Universal Robots URScript: FaiChun_9 Jan_5.script

def Machining1():
  # Default parameters:
  global speed_ms = 0.03
  global speed_rads = 0.75
  global accel_mss = 3
  global accel_radss = 1.2
  global blend_radius_m = 0.0003

  # Add subprograms here
  # Start of main program
  # Program generated by RoboDK v5.6.8 for UR10e on 09/01/2025 17:26:35
  # Using nominal kinematics.
  blend_radius_m = 0.0003
  speed_ms = 0.03
  # set_reference(p[0.325000, -0.070000, 0.000000, 0.000000, 0.000000, 0.000000])
  set_tcp(p[0.000000, 0.000000, 0.252000, 0.000000, 0.000000, 0.000000])
  # Show Tool
  movej([0.354568, -1.073416, -2.632395, -1.006578, 1.570796, 1.925364],accel_radss,speed_rads,0,blend_radius_m)
  movel([0.354568, -1.133460, -2.672124, -0.906805, 1.570796, 1.925364],accel_mss,speed_ms,0,blend_radius_m)
  #SetTool1
  #M_RunCode6
  #3SetRPM60000
  speed_ms = 0.03
  #M_RunCode3
  movel([0.354568, -1.161287, -2.687269, -0.863833, 1.570796, 1.925364],accel_mss,speed_ms,0,blend_radius_m)
  speed_ms = 0.003
  movel([0.354568, -1.168634, -2.690994, -0.852761, 1.570796, 1.925364],accel_mss,speed_ms,0,blend_radius_m)
  speed_ms = 0.007
  movel([0.356966, -1.171496, -2.689722, -0.851171, 1.570796, 1.927762],accel_mss,speed_ms,0,blend_radius_m)
  movel([0.359544, -1.173577, -2.688792, -0.850019, 1.570796, 1.930340],accel_mss,speed_ms,0,blend_radius_m)
  movel([0.362316, -1.174874, -2.688211, -0.849304, 1.570796, 1.933112],accel_mss,speed_ms,0,blend_radius_m)
  movel([0.365281, -1.175393, -2.687978, -0.849019, 1.570796, 1.936077],accel_mss,speed_ms,0,blend_radius_m)
  movel([0.368380, -1.175227, -2.688052, -0.849110, 1.570796, 1.939176],accel_mss,speed_ms,0,blend_radius_m)
  movel([0.371545, -1.174464, -2.688395, -0.849530, 1.570796, 1.942341],accel_mss,speed_ms,0,blend_radius_m)
  movel([0.374787, -1.173102, -2.689005, -0.850282, 1.570796, 1.945583],accel_mss,speed_ms,0,blend_radius_m)
  movel([0.378111, -1.171130, -2.689885, -0.851373, 1.570796, 1.948907],accel_mss,speed_ms,0,blend_radius_m)
  movel([0.363017, -1.184266, -2.683945, -0.844178, 1.570796, 1.933813],accel_mss,speed_ms,0,blend_radius_m)
  movel([0.342026, -1.154782, -2.697027, -0.860579, 1.570796, 1.912822],accel_mss,speed_ms,0,blend_radius_m)
  movel([0.343555, -1.153375, -2.697629, -0.861384, 1.570796, 1.914352],accel_mss,speed_ms,0,blend_radius_m)
  movel([0.347706, -1.150135, -2.699008, -0.863246, 1.570796, 1.918503],accel_mss,speed_ms,0,blend_radius_m)
  movel([0.352300, -1.147640, -2.700062, -0.864686, 1.570796, 1.923096],accel_mss,speed_ms,0,blend_radius_m)
  movel([0.357069, -1.145805, -2.700834, -0.865750, 1.570796, 1.927865],accel_mss,speed_ms,0,blend_radius_m)
  movel([0.361749, -1.144532, -2.701367, -0.866490, 1.570796, 1.932545],accel_mss,speed_ms,0,blend_radius_m)
  movel([0.373963, -1.142426, -2.702246, -0.867717, 1.570796, 1.944759],accel_mss,speed_ms,0,blend_radius_m)
  movel([0.385222, -1.140714, -2.702957, -0.868719, 1.570796, 1.956018],accel_mss,speed_ms,0,blend_radius_m)
  movel([0.389576, -1.139664, -2.703391, -0.869334, 1.570796, 1.960373],accel_mss,speed_ms,0,blend_radius_m)
  movel([0.393934, -1.138139, -2.704021, -0.870229, 1.570796, 1.964730],accel_mss,speed_ms,0,blend_radius_m)
  movel([0.398079, -1.136054, -2.704878, -0.871458, 1.570796, 1.968876],accel_mss,speed_ms,0,blend_radius_m)
  movel([0.401806, -1.133312, -2.705998, -0.873079, 1.570796, 1.972603],accel_mss,speed_ms,0,blend_radius_m)
  movel([0.405715, -1.129228, -2.707653, -0.875508, 1.570796, 1.976512],accel_mss,speed_ms,0,blend_radius_m)
  movel([0.407057, -1.127215, -2.708462, -0.876712, 1.570796, 1.977853],accel_mss,speed_ms,0,blend_radius_m)
  movel([0.407988, -1.125220, -2.709261, -0.877908, 1.570796, 1.978784],accel_mss,speed_ms,0,blend_radius_m)
  movel([0.408720, -1.121628, -2.710690, -0.880072, 1.570796, 1.979516],accel_mss,speed_ms,0,blend_radius_m)
  movel([0.408019, -1.118804, -2.711804, -0.881781, 1.570796, 1.978816],accel_mss,speed_ms,0,blend_radius_m)
  movel([0.406875, -1.117482, -2.712323, -0.882584, 1.570796, 1.977671],accel_mss,speed_ms,0,blend_radius_m)
  movel([0.405474, -1.116991, -2.712516, -0.882883, 1.570796, 1.976271],accel_mss,speed_ms,0,blend_radius_m)
  movel([0.403971, -1.117249, -2.712414, -0.882726, 1.570796, 1.974768],accel_mss,speed_ms,0,blend_radius_m)
  movel([0.402512, -1.118181, -2.712049, -0.882159, 1.570796, 1.973309],accel_mss,speed_ms,0,blend_radius_m)
  movel([0.400903, -1.120447, -2.711157, -0.880785, 1.570796, 1.971699],accel_mss,speed_ms,0,blend_radius_m)
  movel([0.399463, -1.122720, -2.710257, -0.879412, 1.570796, 1.970259],accel_mss,speed_ms,0,blend_radius_m)
  movel([0.397172, -1.125110, -2.709305, -0.877974, 1.570796, 1.967968],accel_mss,speed_ms,0,blend_radius_m)
  movel([0.394069, -1.127271, -2.708440, -0.876678, 1.570796, 1.964865],accel_mss,speed_ms,0,blend_radius_m)
  movel([0.391233, -1.128021, -2.708139, -0.876230, 1.570796, 1.962029],accel_mss,speed_ms,0,blend_radius_m)
  movel([0.388876, -1.127540, -2.708332, -0.876517, 1.570796, 1.959673],accel_mss,speed_ms,0,blend_radius_m)
  movel([0.387215, -1.125994, -2.708952, -0.877443, 1.570796, 1.958012],accel_mss,speed_ms,0,blend_radius_m)
  movel([0.386430, -1.123660, -2.709883, -0.878846, 1.570796, 1.957226],accel_mss,speed_ms,0,blend_radius_m)
  movel([0.386711, -1.120809, -2.711013, -0.880566, 1.570796, 1.957507],accel_mss,speed_ms,0,blend_radius_m)
  movel([0.388136, -1.117739, -2.712222, -0.882428, 1.570796, 1.958932],accel_mss,speed_ms,0,blend_radius_m)
  movel([0.390789, -1.114754, -2.713389, -0.884246, 1.570796, 1.961586],accel_mss,speed_ms,0,blend_radius_m)
  movel([0.393483, -1.112681, -2.714194, -0.885514, 1.570796, 1.964280],accel_mss,speed_ms,0,blend_radius_m)
  movel([0.396144, -1.111333, -2.714716, -0.886340, 1.570796, 1.966940],accel_mss,speed_ms,0,blend_radius_m)
  movel([0.398770, -1.110715, -2.714954, -0.886719, 1.570796, 1.969567],accel_mss,speed_ms,0,blend_radius_m)
  movel([0.401345, -1.110843, -2.714905, -0.886641, 1.570796, 1.972141],accel_mss,speed_ms,0,blend_radius_m)
  movel([0.403780, -1.111624, -2.714603, -0.886161, 1.570796, 1.974576],accel_mss,speed_ms,0,blend_radius_m)
  movel([0.405978, -1.112973, -2.714081, -0.885335, 1.570796, 1.976774],accel_mss,speed_ms,0,blend_radius_m)
  movel([0.409660, -1.117365, -2.712369, -0.882655, 1.570796, 1.980457],accel_mss,speed_ms,0,blend_radius_m)
  movel([0.411296, -1.120837, -2.711002, -0.880549, 1.570796, 1.982092],accel_mss,speed_ms,0,blend_radius_m)
  movel([0.412317, -1.124558, -2.709525, -0.878306, 1.570796, 1.983113],accel_mss,speed_ms,0,blend_radius_m)
  movel([0.412731, -1.128520, -2.707938, -0.875931, 1.570796, 1.983527],accel_mss,speed_ms,0,blend_radius_m)
  movel([0.412549, -1.132708, -2.706243, -0.873438, 1.570796, 1.983345],accel_mss,speed_ms,0,blend_radius_m)
  movel([0.411547, -1.136963, -2.704504, -0.870921, 1.570796, 1.982343],accel_mss,speed_ms,0,blend_radius_m)
  movel([0.409511, -1.141125, -2.702786, -0.868478, 1.570796, 1.980307],accel_mss,speed_ms,0,blend_radius_m)
  movel([0.406444, -1.145198, -2.701088, -0.866103, 1.570796, 1.977240],accel_mss,speed_ms,0,blend_radius_m)
  movel([0.402358, -1.149188, -2.699409, -0.863792, 1.570796, 1.973154],accel_mss,speed_ms,0,blend_radius_m)
  movel([0.398284, -1.152264, -2.698104, -0.862022, 1.570796, 1.969081],accel_mss,speed_ms,0,blend_radius_m)
  movel([0.394157, -1.154540, -2.697131, -0.860718, 1.570796, 1.964954],accel_mss,speed_ms,0,blend_radius_m)
  movel([0.390077, -1.156158, -2.696437, -0.859794, 1.570796, 1.960874],accel_mss,speed_ms,0,blend_radius_m)
  movel([0.386157, -1.157252, -2.695966, -0.859171, 1.570796, 1.956954],accel_mss,speed_ms,0,blend_radius_m)
  movel([0.376830, -1.158761, -2.695314, -0.858314, 1.570796, 1.947626],accel_mss,speed_ms,0,blend_radius_m)
  movel([0.367992, -1.160305, -2.694646, -0.857439, 1.570796, 1.938788],accel_mss,speed_ms,0,blend_radius_m)
  movel([0.364425, -1.161338, -2.694196, -0.856855, 1.570796, 1.935222],accel_mss,speed_ms,0,blend_radius_m)
  movel([0.360783, -1.162831, -2.693545, -0.856012, 1.570796, 1.931580],accel_mss,speed_ms,0,blend_radius_m)
  movel([0.357192, -1.164865, -2.692655, -0.854869, 1.570796, 1.927988],accel_mss,speed_ms,0,blend_radius_m)
  movel([0.353786, -1.167525, -2.691484, -0.853380, 1.570796, 1.924582],accel_mss,speed_ms,0,blend_radius_m)
  movel([0.354568, -1.168634, -2.690994, -0.852761, 1.570796, 1.925364],accel_mss,speed_ms,0,blend_radius_m)
  speed_ms = 0.003
  movel([0.354568, -1.161287, -2.687269, -0.863833, 1.570796, 1.925364],accel_mss,speed_ms,0,blend_radius_m)
  speed_ms = 0.03
  movel([0.354568, -1.133460, -2.672124, -0.906805, 1.570796, 1.925364],accel_mss,speed_ms,0,blend_radius_m)
  #M_RunCode9
  movel([0.379678, -1.157713, -2.661566, -0.893110, 1.570796, 1.950474],accel_mss,speed_ms,0,blend_radius_m)
  #M_RunCode3
  movel([0.379678, -1.185401, -2.676392, -0.850596, 1.570796, 1.950474],accel_mss,speed_ms,0,blend_radius_m)
  speed_ms = 0.003
  movel([0.379678, -1.192696, -2.680036, -0.839657, 1.570796, 1.950474],accel_mss,speed_ms,0,blend_radius_m)
  speed_ms = 0.007
  movel([0.387460, -1.185010, -2.683603, -0.843776, 1.570796, 1.958256],accel_mss,speed_ms,0,blend_radius_m)
  movel([0.399155, -1.174764, -2.688260, -0.849365, 1.570796, 1.969951],accel_mss,speed_ms,0,blend_radius_m)
  movel([0.411336, -1.164890, -2.692644, -0.854855, 1.570796, 1.982132],accel_mss,speed_ms,0,blend_radius_m)
  movel([0.420366, -1.158451, -2.695449, -0.858490, 1.570796, 1.991162],accel_mss,speed_ms,0,blend_radius_m)
  movel([0.423713, -1.156585, -2.696253, -0.859551, 1.570796, 1.994510],accel_mss,speed_ms,0,blend_radius_m)
  movel([0.426343, -1.155682, -2.696642, -0.860066, 1.570796, 1.997139],accel_mss,speed_ms,0,blend_radius_m)
  movel([0.428246, -1.155744, -2.696615, -0.860030, 1.570796, 1.999042],accel_mss,speed_ms,0,blend_radius_m)
  movel([0.429420, -1.156775, -2.696172, -0.859443, 1.570796, 2.000216],accel_mss,speed_ms,0,blend_radius_m)
  movel([0.429733, -1.158510, -2.695423, -0.858456, 1.570796, 2.000529],accel_mss,speed_ms,0,blend_radius_m)
  movel([0.429055, -1.160703, -2.694472, -0.857213, 1.570796, 1.999851],accel_mss,speed_ms,0,blend_radius_m)
  movel([0.427394, -1.163343, -2.693322, -0.855724, 1.570796, 1.998190],accel_mss,speed_ms,0,blend_radius_m)
  movel([0.424759, -1.166426, -2.691969, -0.853994, 1.570796, 1.995555],accel_mss,speed_ms,0,blend_radius_m)
  movel([0.416644, -1.174214, -2.688507, -0.849668, 1.570796, 1.987440],accel_mss,speed_ms,0,blend_radius_m)
  movel([0.404851, -1.184338, -2.683912, -0.844139, 1.570796, 1.975647],accel_mss,speed_ms,0,blend_radius_m)
  movel([0.392963, -1.193873, -2.679484, -0.839032, 1.570796, 1.963760],accel_mss,speed_ms,0,blend_radius_m)
  movel([0.384351, -1.200009, -2.676582, -0.835798, 1.570796, 1.955147],accel_mss,speed_ms,0,blend_radius_m)
  movel([0.381176, -1.201791, -2.675731, -0.834866, 1.570796, 1.951973],accel_mss,speed_ms,0,blend_radius_m)
  movel([0.378665, -1.202681, -2.675305, -0.834403, 1.570796, 1.949461],accel_mss,speed_ms,0,blend_radius_m)
  movel([0.376810, -1.202676, -2.675308, -0.834405, 1.570796, 1.947607],accel_mss,speed_ms,0,blend_radius_m)
  movel([0.375605, -1.201780, -2.675737, -0.834872, 1.570796, 1.946401],accel_mss,speed_ms,0,blend_radius_m)
  movel([0.375198, -1.200206, -2.676488, -0.835695, 1.570796, 1.945994],accel_mss,speed_ms,0,blend_radius_m)
  movel([0.375736, -1.198170, -2.677456, -0.836763, 1.570796, 1.946532],accel_mss,speed_ms,0,blend_radius_m)
  movel([0.377227, -1.195668, -2.678639, -0.838082, 1.570796, 1.948024],accel_mss,speed_ms,0,blend_radius_m)
  movel([0.379678, -1.192696, -2.680036, -0.839657, 1.570796, 1.950474],accel_mss,speed_ms,0,blend_radius_m)
  speed_ms = 0.003
  movel([0.379678, -1.185401, -2.676392, -0.850596, 1.570796, 1.950474],accel_mss,speed_ms,0,blend_radius_m)
  speed_ms = 0.03
  movel([0.379678, -1.157713, -2.661566, -0.893110, 1.570796, 1.950474],accel_mss,speed_ms,0,blend_radius_m)
  #M_RunCode9
  movel([0.372229, -1.160949, -2.660112, -0.891327, 1.570796, 1.943026],accel_mss,speed_ms,0,blend_radius_m)
  #M_RunCode3
  movel([0.372229, -1.188615, -2.674896, -0.848878, 1.570796, 1.943026],accel_mss,speed_ms,0,blend_radius_m)
  speed_ms = 0.003
  movel([0.372229, -1.195902, -2.678528, -0.837958, 1.570796, 1.943026],accel_mss,speed_ms,0,blend_radius_m)
  speed_ms = 0.007
  movel([0.372519, -1.193032, -2.679878, -0.839479, 1.570796, 1.943316],accel_mss,speed_ms,0,blend_radius_m)
  movel([0.373292, -1.189945, -2.681319, -0.841124, 1.570796, 1.944089],accel_mss,speed_ms,0,blend_radius_m)
  movel([0.374568, -1.186684, -2.682831, -0.842874, 1.570796, 1.945364],accel_mss,speed_ms,0,blend_radius_m)
  movel([0.376355, -1.183240, -2.684415, -0.844734, 1.570796, 1.947151],accel_mss,speed_ms,0,blend_radius_m)
  movel([0.378653, -1.179619, -2.686067, -0.846703, 1.570796, 1.949450],accel_mss,speed_ms,0,blend_radius_m)
  movel([0.381456, -1.175876, -2.687760, -0.848753, 1.570796, 1.952252],accel_mss,speed_ms,0,blend_radius_m)
  movel([0.384749, -1.172089, -2.689458, -0.850842, 1.570796, 1.955546],accel_mss,speed_ms,0,blend_radius_m)
  movel([0.388543, -1.168254, -2.691162, -0.852973, 1.570796, 1.959339],accel_mss,speed_ms,0,blend_radius_m)
  movel([0.392836, -1.164375, -2.692870, -0.855144, 1.570796, 1.963633],accel_mss,speed_ms,0,blend_radius_m)
  movel([0.397312, -1.160734, -2.694459, -0.857196, 1.570796, 1.968109],accel_mss,speed_ms,0,blend_radius_m)
  movel([0.401640, -1.157615, -2.695810, -0.858965, 1.570796, 1.972436],accel_mss,speed_ms,0,blend_radius_m)
  movel([0.405819, -1.155020, -2.696926, -0.860443, 1.570796, 1.976615],accel_mss,speed_ms,0,blend_radius_m)
  movel([0.409833, -1.152965, -2.697805, -0.861619, 1.570796, 1.980629],accel_mss,speed_ms,0,blend_radius_m)
  movel([0.413614, -1.151451, -2.698450, -0.862489, 1.570796, 1.984410],accel_mss,speed_ms,0,blend_radius_m)
  movel([0.417092, -1.150479, -2.698862, -0.863048, 1.570796, 1.987889],accel_mss,speed_ms,0,blend_radius_m)
  movel([0.420254, -1.150059, -2.699040, -0.863290, 1.570796, 1.991051],accel_mss,speed_ms,0,blend_radius_m)
  movel([0.423104, -1.150185, -2.698987, -0.863217, 1.570796, 1.993900],accel_mss,speed_ms,0,blend_radius_m)
  movel([0.425609, -1.150820, -2.698717, -0.862851, 1.570796, 1.996406],accel_mss,speed_ms,0,blend_radius_m)
  movel([0.427747, -1.151930, -2.698246, -0.862214, 1.570796, 1.998543],accel_mss,speed_ms,0,blend_radius_m)
  movel([0.429513, -1.153503, -2.697575, -0.861311, 1.570796, 2.000309],accel_mss,speed_ms,0,blend_radius_m)
  movel([0.430906, -1.155546, -2.696700, -0.860143, 1.570796, 2.001703],accel_mss,speed_ms,0,blend_radius_m)
  movel([0.431874, -1.157931, -2.695673, -0.858785, 1.570796, 2.002670],accel_mss,speed_ms,0,blend_radius_m)
  movel([0.432358, -1.160544, -2.694541, -0.857303, 1.570796, 2.003155],accel_mss,speed_ms,0,blend_radius_m)
  movel([0.432364, -1.163381, -2.693305, -0.855703, 1.570796, 2.003160],accel_mss,speed_ms,0,blend_radius_m)
  movel([0.431892, -1.166435, -2.691965, -0.853989, 1.570796, 2.002688],accel_mss,speed_ms,0,blend_radius_m)
  movel([0.430933, -1.169665, -2.690537, -0.852187, 1.570796, 2.001729],accel_mss,speed_ms,0,blend_radius_m)
  movel([0.429473, -1.173023, -2.689040, -0.850325, 1.570796, 2.000269],accel_mss,speed_ms,0,blend_radius_m)
  movel([0.427521, -1.176505, -2.687476, -0.848407, 1.570796, 1.998318],accel_mss,speed_ms,0,blend_radius_m)
  movel([0.425078, -1.180116, -2.685842, -0.846432, 1.570796, 1.995874],accel_mss,speed_ms,0,blend_radius_m)
  movel([0.422172, -1.183774, -2.684170, -0.844444, 1.570796, 1.992968],accel_mss,speed_ms,0,blend_radius_m)
  movel([0.418832, -1.187414, -2.682494, -0.842481, 1.570796, 1.989629],accel_mss,speed_ms,0,blend_radius_m)
  movel([0.415055, -1.191041, -2.680809, -0.840539, 1.570796, 1.985852],accel_mss,speed_ms,0,blend_radius_m)
  movel([0.410849, -1.194652, -2.679117, -0.838619, 1.570796, 1.981646],accel_mss,speed_ms,0,blend_radius_m)
  movel([0.406521, -1.198006, -2.677534, -0.836850, 1.570796, 1.977317],accel_mss,speed_ms,0,blend_radius_m)
  movel([0.402383, -1.200845, -2.676183, -0.835360, 1.570796, 1.973179],accel_mss,speed_ms,0,blend_radius_m)
  movel([0.398419, -1.203189, -2.675062, -0.834138, 1.570796, 1.969215],accel_mss,speed_ms,0,blend_radius_m)
  movel([0.394629, -1.205036, -2.674174, -0.833179, 1.570796, 1.965426],accel_mss,speed_ms,0,blend_radius_m)
  movel([0.391062, -1.206401, -2.673515, -0.832473, 1.570796, 1.961858],accel_mss,speed_ms,0,blend_radius_m)
  movel([0.387772, -1.207286, -2.673087, -0.832016, 1.570796, 1.958568],accel_mss,speed_ms,0,blend_radius_m)
  movel([0.384754, -1.207698, -2.672887, -0.831804, 1.570796, 1.955550],accel_mss,speed_ms,0,blend_radius_m)
  movel([0.382004, -1.207633, -2.672919, -0.831838, 1.570796, 1.952800],accel_mss,speed_ms,0,blend_radius_m)
  movel([0.379552, -1.207117, -2.673169, -0.832104, 1.570796, 1.950348],accel_mss,speed_ms,0,blend_radius_m)
  movel([0.377425, -1.206179, -2.673622, -0.832588, 1.570796, 1.948222],accel_mss,speed_ms,0,blend_radius_m)
  movel([0.375621, -1.204815, -2.674280, -0.833294, 1.570796, 1.946417],accel_mss,speed_ms,0,blend_radius_m)
  movel([0.374138, -1.203022, -2.675142, -0.834225, 1.570796, 1.944934],accel_mss,speed_ms,0,blend_radius_m)
  movel([0.373043, -1.200893, -2.676161, -0.835336, 1.570796, 1.943839],accel_mss,speed_ms,0,blend_radius_m)
  movel([0.372405, -1.198522, -2.677289, -0.836578, 1.570796, 1.943201],accel_mss,speed_ms,0,blend_radius_m)
  movel([0.372229, -1.195902, -2.678528, -0.837958, 1.570796, 1.943026],accel_mss,speed_ms,0,blend_radius_m)
  speed_ms = 0.003
  movel([0.372229, -1.188615, -2.674896, -0.848878, 1.570796, 1.943026],accel_mss,speed_ms,0,blend_radius_m)
  speed_ms = 0.03
  movel([0.372229, -1.160949, -2.660112, -0.891327, 1.570796, 1.943026],accel_mss,speed_ms,0,blend_radius_m)
  #M_RunCode9
  movel([0.502532, -1.419663, -2.504293, -0.788433, 1.570796, 2.073328],accel_mss,speed_ms,0,blend_radius_m)
  #M_RunCode3
  movel([0.502532, -1.443463, -2.515724, -0.753202, 1.570796, 2.073328],accel_mss,speed_ms,0,blend_radius_m)
  speed_ms = 0.003
  movel([0.502532, -1.449619, -2.518509, -0.744260, 1.570796, 2.073328],accel_mss,speed_ms,0,blend_radius_m)
  speed_ms = 0.007
  movel([0.503681, -1.448967, -2.519037, -0.744386, 1.570796, 2.074477],accel_mss,speed_ms,0,blend_radius_m)
  movel([0.506715, -1.447598, -2.520141, -0.744650, 1.570796, 2.077511],accel_mss,speed_ms,0,blend_radius_m)
  movel([0.509926, -1.446841, -2.520750, -0.744798, 1.570796, 2.080722],accel_mss,speed_ms,0,blend_radius_m)
  movel([0.513159, -1.446571, -2.520967, -0.744851, 1.570796, 2.083955],accel_mss,speed_ms,0,blend_radius_m)
  movel([0.516261, -1.446673, -2.520885, -0.744831, 1.570796, 2.087058],accel_mss,speed_ms,0,blend_radius_m)
  movel([0.524203, -1.447750, -2.520018, -0.744621, 1.570796, 2.094999],accel_mss,speed_ms,0,blend_radius_m)
  movel([0.531487, -1.448876, -2.519110, -0.744403, 1.570796, 2.102283],accel_mss,speed_ms,0,blend_radius_m)
  movel([0.534346, -1.449044, -2.518974, -0.744371, 1.570796, 2.105142],accel_mss,speed_ms,0,blend_radius_m)
  movel([0.537257, -1.448890, -2.519099, -0.744400, 1.570796, 2.108054],accel_mss,speed_ms,0,blend_radius_m)
  movel([0.540096, -1.448313, -2.519564, -0.744512, 1.570796, 2.110892],accel_mss,speed_ms,0,blend_radius_m)
  movel([0.542736, -1.447217, -2.520447, -0.744724, 1.570796, 2.113533],accel_mss,speed_ms,0,blend_radius_m)
  movel([0.545632, -1.445261, -2.522019, -0.745109, 1.570796, 2.116429],accel_mss,speed_ms,0,blend_radius_m)
  movel([0.546690, -1.444183, -2.522883, -0.745323, 1.570796, 2.117486],accel_mss,speed_ms,0,blend_radius_m)
  movel([0.547489, -1.443035, -2.523801, -0.745553, 1.570796, 2.118285],accel_mss,speed_ms,0,blend_radius_m)
  movel([0.548333, -1.440787, -2.525592, -0.746010, 1.570796, 2.119129],accel_mss,speed_ms,0,blend_radius_m)
  movel([0.548201, -1.438765, -2.527197, -0.746427, 1.570796, 2.118997],accel_mss,speed_ms,0,blend_radius_m)
  movel([0.547632, -1.437654, -2.528076, -0.746659, 1.570796, 2.118428],accel_mss,speed_ms,0,blend_radius_m)
  movel([0.546815, -1.437041, -2.528560, -0.746788, 1.570796, 2.117611],accel_mss,speed_ms,0,blend_radius_m)
  movel([0.545850, -1.436910, -2.528664, -0.746815, 1.570796, 2.116646],accel_mss,speed_ms,0,blend_radius_m)
  movel([0.544842, -1.437235, -2.528407, -0.746747, 1.570796, 2.115638],accel_mss,speed_ms,0,blend_radius_m)
  movel([0.543588, -1.438420, -2.527470, -0.746499, 1.570796, 2.114384],accel_mss,speed_ms,0,blend_radius_m)
  movel([0.542440, -1.439645, -2.526499, -0.746245, 1.570796, 2.113236],accel_mss,speed_ms,0,blend_radius_m)
  movel([0.540743, -1.440783, -2.525595, -0.746011, 1.570796, 2.111539],accel_mss,speed_ms,0,blend_radius_m)
  movel([0.538563, -1.441600, -2.524945, -0.745844, 1.570796, 2.109360],accel_mss,speed_ms,0,blend_radius_m)
  movel([0.536708, -1.441527, -2.525003, -0.745859, 1.570796, 2.107504],accel_mss,speed_ms,0,blend_radius_m)
  movel([0.535289, -1.440723, -2.525643, -0.746023, 1.570796, 2.106086],accel_mss,speed_ms,0,blend_radius_m)
  movel([0.534426, -1.439342, -2.526740, -0.746307, 1.570796, 2.105222],accel_mss,speed_ms,0,blend_radius_m)
  movel([0.534206, -1.437610, -2.528111, -0.746668, 1.570796, 2.105002],accel_mss,speed_ms,0,blend_radius_m)
  movel([0.534705, -1.435753, -2.529576, -0.747060, 1.570796, 2.105502],accel_mss,speed_ms,0,blend_radius_m)
  movel([0.535944, -1.433987, -2.530964, -0.747438, 1.570796, 2.106741],accel_mss,speed_ms,0,blend_radius_m)
  movel([0.537934, -1.432538, -2.532100, -0.747751, 1.570796, 2.108730],accel_mss,speed_ms,0,blend_radius_m)
  movel([0.539842, -1.431708, -2.532749, -0.747932, 1.570796, 2.110639],accel_mss,speed_ms,0,blend_radius_m)
  movel([0.541646, -1.431359, -2.533022, -0.748008, 1.570796, 2.112443],accel_mss,speed_ms,0,blend_radius_m)
  movel([0.543341, -1.431492, -2.532918, -0.747979, 1.570796, 2.114137],accel_mss,speed_ms,0,blend_radius_m)
  movel([0.544925, -1.432107, -2.532437, -0.747845, 1.570796, 2.115721],accel_mss,speed_ms,0,blend_radius_m)
  movel([0.546349, -1.433124, -2.531641, -0.747624, 1.570796, 2.117145],accel_mss,speed_ms,0,blend_radius_m)
  movel([0.547567, -1.434472, -2.530584, -0.747334, 1.570796, 2.118363],accel_mss,speed_ms,0,blend_radius_m)
  movel([0.549380, -1.438137, -2.527694, -0.746558, 1.570796, 2.120176],accel_mss,speed_ms,0,blend_radius_m)
  movel([0.550024, -1.440778, -2.525599, -0.746012, 1.570796, 2.120821],accel_mss,speed_ms,0,blend_radius_m)
  movel([0.550264, -1.443459, -2.523462, -0.745468, 1.570796, 2.121061],accel_mss,speed_ms,0,blend_radius_m)
  movel([0.550102, -1.446181, -2.521280, -0.744927, 1.570796, 2.120899],accel_mss,speed_ms,0,blend_radius_m)
  movel([0.549541, -1.448944, -2.519055, -0.744390, 1.570796, 2.120337],accel_mss,speed_ms,0,blend_radius_m)
  movel([0.548461, -1.451593, -2.516910, -0.743886, 1.570796, 2.119258],accel_mss,speed_ms,0,blend_radius_m)
  movel([0.546732, -1.453987, -2.514963, -0.743439, 1.570796, 2.117528],accel_mss,speed_ms,0,blend_radius_m)
  movel([0.544360, -1.456125, -2.513216, -0.743048, 1.570796, 2.115156],accel_mss,speed_ms,0,blend_radius_m)
  movel([0.541346, -1.458015, -2.511666, -0.742708, 1.570796, 2.112142],accel_mss,speed_ms,0,blend_radius_m)
  movel([0.538430, -1.459300, -2.510609, -0.742480, 1.570796, 2.109226],accel_mss,speed_ms,0,blend_radius_m)
  movel([0.535563, -1.460034, -2.510004, -0.742351, 1.570796, 2.106359],accel_mss,speed_ms,0,blend_radius_m)
  movel([0.532795, -1.460332, -2.509758, -0.742299, 1.570796, 2.103591],accel_mss,speed_ms,0,blend_radius_m)
  movel([0.530186, -1.460301, -2.509784, -0.742304, 1.570796, 2.100982],accel_mss,speed_ms,0,blend_radius_m)
  movel([0.524093, -1.459478, -2.510462, -0.742449, 1.570796, 2.094889],accel_mss,speed_ms,0,blend_radius_m)
  movel([0.518303, -1.458764, -2.511050, -0.742575, 1.570796, 2.089099],accel_mss,speed_ms,0,blend_radius_m)
  movel([0.515911, -1.458756, -2.511056, -0.742576, 1.570796, 2.086707],accel_mss,speed_ms,0,blend_radius_m)
  movel([0.513417, -1.459046, -2.510818, -0.742525, 1.570796, 2.084213],accel_mss,speed_ms,0,blend_radius_m)
  movel([0.510883, -1.459724, -2.510260, -0.742405, 1.570796, 2.081680],accel_mss,speed_ms,0,blend_radius_m)
  movel([0.508387, -1.460872, -2.509313, -0.742205, 1.570796, 2.079183],accel_mss,speed_ms,0,blend_radius_m)
  movel([0.508747, -1.461799, -2.508546, -0.742044, 1.570796, 2.079544],accel_mss,speed_ms,0,blend_radius_m)
  movel([0.509923, -1.464268, -2.506499, -0.741623, 1.570796, 2.080720],accel_mss,speed_ms,0,blend_radius_m)
  movel([0.511316, -1.466229, -2.504866, -0.741295, 1.570796, 2.082112],accel_mss,speed_ms,0,blend_radius_m)
  movel([0.512928, -1.467681, -2.503653, -0.741056, 1.570796, 2.083724],accel_mss,speed_ms,0,blend_radius_m)
  movel([0.514763, -1.468630, -2.502858, -0.740901, 1.570796, 2.085560],accel_mss,speed_ms,0,blend_radius_m)
  movel([0.516763, -1.469129, -2.502439, -0.740820, 1.570796, 2.087560],accel_mss,speed_ms,0,blend_radius_m)
  movel([0.518878, -1.469227, -2.502357, -0.740805, 1.570796, 2.089674],accel_mss,speed_ms,0,blend_radius_m)
  movel([0.521111, -1.468926, -2.502610, -0.740853, 1.570796, 2.091907],accel_mss,speed_ms,0,blend_radius_m)
  movel([0.523464, -1.468222, -2.503200, -0.740967, 1.570796, 2.094261],accel_mss,speed_ms,0,blend_radius_m)
  movel([0.512242, -1.474339, -2.498048, -0.740001, 1.570796, 2.083038],accel_mss,speed_ms,0,blend_radius_m)
  movel([0.502532, -1.449619, -2.518509, -0.744260, 1.570796, 2.073328],accel_mss,speed_ms,0,blend_radius_m)
  speed_ms = 0.003
  movel([0.502532, -1.443463, -2.515724, -0.753202, 1.570796, 2.073328],accel_mss,speed_ms,0,blend_radius_m)
  speed_ms = 0.03
  movel([0.502532, -1.419663, -2.504293, -0.788433, 1.570796, 2.073328],accel_mss,speed_ms,0,blend_radius_m)
  #M_RunCode9
  movel([0.520386, -1.444284, -2.484836, -0.783269, 1.570796, 2.091182],accel_mss,speed_ms,0,blend_radius_m)
  #M_RunCode3
  movel([0.520386, -1.467574, -2.495971, -0.748844, 1.570796, 2.091182],accel_mss,speed_ms,0,blend_radius_m)
  speed_ms = 0.003
  movel([0.520386, -1.473591, -2.498682, -0.740116, 1.570796, 2.091182],accel_mss,speed_ms,0,blend_radius_m)
  speed_ms = 0.007
  movel([0.522489, -1.472799, -2.499351, -0.740239, 1.570796, 2.093285],accel_mss,speed_ms,0,blend_radius_m)
  movel([0.524314, -1.472851, -2.499307, -0.740231, 1.570796, 2.095110],accel_mss,speed_ms,0,blend_radius_m)
  movel([0.525722, -1.473608, -2.498667, -0.740114, 1.570796, 2.096518],accel_mss,speed_ms,0,blend_radius_m)
  movel([0.526574, -1.474922, -2.497555, -0.739912, 1.570796, 2.097370],accel_mss,speed_ms,0,blend_radius_m)
  movel([0.526791, -1.476572, -2.496153, -0.739663, 1.570796, 2.097588],accel_mss,speed_ms,0,blend_radius_m)
  movel([0.526305, -1.478339, -2.494649, -0.739401, 1.570796, 2.097101],accel_mss,speed_ms,0,blend_radius_m)
  movel([0.525120, -1.480001, -2.493229, -0.739159, 1.570796, 2.095916],accel_mss,speed_ms,0,blend_radius_m)
  movel([0.523245, -1.481345, -2.492077, -0.738967, 1.570796, 2.094042],accel_mss,speed_ms,0,blend_radius_m)
  movel([0.521515, -1.482061, -2.491462, -0.738865, 1.570796, 2.092311],accel_mss,speed_ms,0,blend_radius_m)
  movel([0.520091, -1.482250, -2.491300, -0.738839, 1.570796, 2.090887],accel_mss,speed_ms,0,blend_radius_m)
  movel([0.518624, -1.482555, -2.491038, -0.738796, 1.570796, 2.089421],accel_mss,speed_ms,0,blend_radius_m)
  movel([0.517799, -1.483212, -2.490473, -0.738704, 1.570796, 2.088595],accel_mss,speed_ms,0,blend_radius_m)
  movel([0.517265, -1.484139, -2.489674, -0.738576, 1.570796, 2.088062],accel_mss,speed_ms,0,blend_radius_m)
  movel([0.517061, -1.485175, -2.488781, -0.738434, 1.570796, 2.087857],accel_mss,speed_ms,0,blend_radius_m)
  movel([0.517236, -1.486156, -2.487933, -0.738301, 1.570796, 2.088032],accel_mss,speed_ms,0,blend_radius_m)
  movel([0.517843, -1.487249, -2.486986, -0.738154, 1.570796, 2.088640],accel_mss,speed_ms,0,blend_radius_m)
  movel([0.518742, -1.488058, -2.486284, -0.738047, 1.570796, 2.089539],accel_mss,speed_ms,0,blend_radius_m)
  movel([0.519931, -1.488587, -2.485824, -0.737978, 1.570796, 2.090728],accel_mss,speed_ms,0,blend_radius_m)
  movel([0.521411, -1.488838, -2.485606, -0.737945, 1.570796, 2.092207],accel_mss,speed_ms,0,blend_radius_m)
  movel([0.523094, -1.488797, -2.485642, -0.737951, 1.570796, 2.093890],accel_mss,speed_ms,0,blend_radius_m)
  movel([0.524895, -1.488450, -2.485943, -0.737996, 1.570796, 2.095692],accel_mss,speed_ms,0,blend_radius_m)
  movel([0.526817, -1.487796, -2.486511, -0.738082, 1.570796, 2.097614],accel_mss,speed_ms,0,blend_radius_m)
  movel([0.528859, -1.486838, -2.487342, -0.738209, 1.570796, 2.099656],accel_mss,speed_ms,0,blend_radius_m)
  movel([0.532082, -1.484699, -2.489191, -0.738499, 1.570796, 2.102878],accel_mss,speed_ms,0,blend_radius_m)
  movel([0.534713, -1.481997, -2.491517, -0.738874, 1.570796, 2.105509],accel_mss,speed_ms,0,blend_radius_m)
  movel([0.535775, -1.480445, -2.492849, -0.739095, 1.570796, 2.106572],accel_mss,speed_ms,0,blend_radius_m)
  movel([0.536623, -1.478770, -2.494281, -0.739338, 1.570796, 2.107420],accel_mss,speed_ms,0,blend_radius_m)
  movel([0.537680, -1.475052, -2.497444, -0.739893, 1.570796, 2.108477],accel_mss,speed_ms,0,blend_radius_m)
  movel([0.537768, -1.470939, -2.500919, -0.740531, 1.570796, 2.108564],accel_mss,speed_ms,0,blend_radius_m)
  movel([0.536756, -1.466539, -2.504607, -0.741243, 1.570796, 2.107552],accel_mss,speed_ms,0,blend_radius_m)
  movel([0.554264, -1.457346, -2.512215, -0.742828, 1.570796, 2.125060],accel_mss,speed_ms,0,blend_radius_m)
  movel([0.560234, -1.476474, -2.496237, -0.739678, 1.570796, 2.131030],accel_mss,speed_ms,0,blend_radius_m)
  movel([0.549016, -1.482190, -2.491352, -0.738847, 1.570796, 2.119813],accel_mss,speed_ms,0,blend_radius_m)
  movel([0.551456, -1.480107, -2.493138, -0.739144, 1.570796, 2.122253],accel_mss,speed_ms,0,blend_radius_m)
  movel([0.553474, -1.477547, -2.495324, -0.739518, 1.570796, 2.124270],accel_mss,speed_ms,0,blend_radius_m)
  movel([0.554963, -1.474628, -2.497804, -0.739957, 1.570796, 2.125759],accel_mss,speed_ms,0,blend_radius_m)
  movel([0.555816, -1.471477, -2.500466, -0.740446, 1.570796, 2.126612],accel_mss,speed_ms,0,blend_radius_m)
  movel([0.555965, -1.468214, -2.503206, -0.740969, 1.570796, 2.126762],accel_mss,speed_ms,0,blend_radius_m)
  movel([0.555338, -1.464970, -2.505915, -0.741504, 1.570796, 2.126134],accel_mss,speed_ms,0,blend_radius_m)
  movel([0.542493, -1.471640, -2.500329, -0.740420, 1.570796, 2.113289],accel_mss,speed_ms,0,blend_radius_m)
  movel([0.543387, -1.475544, -2.497027, -0.739818, 1.570796, 2.114183],accel_mss,speed_ms,0,blend_radius_m)
  movel([0.543518, -1.479641, -2.493536, -0.739211, 1.570796, 2.114314],accel_mss,speed_ms,0,blend_radius_m)
  movel([0.542781, -1.483707, -2.490047, -0.738635, 1.570796, 2.113577],accel_mss,speed_ms,0,blend_radius_m)
  movel([0.542044, -1.485647, -2.488372, -0.738369, 1.570796, 2.112841],accel_mss,speed_ms,0,blend_radius_m)
  movel([0.541062, -1.487526, -2.486746, -0.738118, 1.570796, 2.111859],accel_mss,speed_ms,0,blend_radius_m)
  movel([0.539817, -1.489287, -2.485216, -0.737887, 1.570796, 2.110614],accel_mss,speed_ms,0,blend_radius_m)
  movel([0.538291, -1.490874, -2.483832, -0.737683, 1.570796, 2.109087],accel_mss,speed_ms,0,blend_radius_m)
  movel([0.536486, -1.492288, -2.482597, -0.737504, 1.570796, 2.107282],accel_mss,speed_ms,0,blend_radius_m)
  movel([0.534398, -1.493535, -2.481505, -0.737350, 1.570796, 2.105194],accel_mss,speed_ms,0,blend_radius_m)
  movel([0.532220, -1.494525, -2.480635, -0.737228, 1.570796, 2.103017],accel_mss,speed_ms,0,blend_radius_m)
  movel([0.530142, -1.495171, -2.480068, -0.737150, 1.570796, 2.100938],accel_mss,speed_ms,0,blend_radius_m)
  movel([0.528159, -1.495475, -2.479801, -0.737114, 1.570796, 2.098955],accel_mss,speed_ms,0,blend_radius_m)
  movel([0.526270, -1.495438, -2.479833, -0.737118, 1.570796, 2.097067],accel_mss,speed_ms,0,blend_radius_m)
  movel([0.522880, -1.494557, -2.480607, -0.737225, 1.570796, 2.093677],accel_mss,speed_ms,0,blend_radius_m)
  movel([0.520066, -1.492746, -2.482196, -0.737447, 1.570796, 2.090862],accel_mss,speed_ms,0,blend_radius_m)
  movel([0.517868, -1.490233, -2.484392, -0.737765, 1.570796, 2.088664],accel_mss,speed_ms,0,blend_radius_m)
  movel([0.516324, -1.487254, -2.486981, -0.738154, 1.570796, 2.087120],accel_mss,speed_ms,0,blend_radius_m)
  movel([0.515726, -1.484957, -2.488969, -0.738463, 1.570796, 2.086522],accel_mss,speed_ms,0,blend_radius_m)
  movel([0.515564, -1.482385, -2.491184, -0.738820, 1.570796, 2.086361],accel_mss,speed_ms,0,blend_radius_m)
  movel([0.515904, -1.479753, -2.493441, -0.739195, 1.570796, 2.086700],accel_mss,speed_ms,0,blend_radius_m)
  movel([0.516813, -1.477278, -2.495553, -0.739558, 1.570796, 2.087609],accel_mss,speed_ms,0,blend_radius_m)
  movel([0.518302, -1.475158, -2.497355, -0.739877, 1.570796, 2.089099],accel_mss,speed_ms,0,blend_radius_m)
  movel([0.520386, -1.473591, -2.498682, -0.740116, 1.570796, 2.091182],accel_mss,speed_ms,0,blend_radius_m)
  speed_ms = 0.003
  movel([0.520386, -1.467574, -2.495971, -0.748844, 1.570796, 2.091182],accel_mss,speed_ms,0,blend_radius_m)
  speed_ms = 0.03
  movel([0.520386, -1.444284, -2.484836, -0.783269, 1.570796, 2.091182],accel_mss,speed_ms,0,blend_radius_m)
  #M_RunCode9
  movel([0.530140, -1.341533, -2.560339, -0.810516, 1.570796, 2.100936],accel_mss,speed_ms,0,blend_radius_m)
  #M_RunCode3
  movel([0.530140, -1.366842, -2.572748, -0.772799, 1.570796, 2.100936],accel_mss,speed_ms,0,blend_radius_m)
  speed_ms = 0.003
  movel([0.530140, -1.373419, -2.575779, -0.763191, 1.570796, 2.100936],accel_mss,speed_ms,0,blend_radius_m)
  speed_ms = 0.007
  movel([0.526555, -1.374010, -2.575367, -0.763012, 1.570796, 2.097352],accel_mss,speed_ms,0,blend_radius_m)
  movel([0.523091, -1.373873, -2.575462, -0.763053, 1.570796, 2.093887],accel_mss,speed_ms,0,blend_radius_m)
  movel([0.519810, -1.373139, -2.575973, -0.763277, 1.570796, 2.090607],accel_mss,speed_ms,0,blend_radius_m)
  movel([0.516789, -1.371928, -2.576814, -0.763646, 1.570796, 2.087585],accel_mss,speed_ms,0,blend_radius_m)
  movel([0.514105, -1.370358, -2.577902, -0.764129, 1.570796, 2.084901],accel_mss,speed_ms,0,blend_radius_m)
  movel([0.516210, -1.366248, -2.580732, -0.765409, 1.570796, 2.087007],accel_mss,speed_ms,0,blend_radius_m)
  movel([0.519512, -1.361869, -2.583721, -0.766799, 1.570796, 2.090309],accel_mss,speed_ms,0,blend_radius_m)
  movel([0.523673, -1.357616, -2.586598, -0.768175, 1.570796, 2.094469],accel_mss,speed_ms,0,blend_radius_m)
  movel([0.528331, -1.353900, -2.589091, -0.769398, 1.570796, 2.099127],accel_mss,speed_ms,0,blend_radius_m)
  movel([0.533122, -1.351134, -2.590934, -0.770321, 1.570796, 2.103918],accel_mss,speed_ms,0,blend_radius_m)
  movel([0.535444, -1.350240, -2.591528, -0.770621, 1.570796, 2.106241],accel_mss,speed_ms,0,blend_radius_m)
  movel([0.537660, -1.349738, -2.591860, -0.770790, 1.570796, 2.108456],accel_mss,speed_ms,0,blend_radius_m)
  movel([0.539711, -1.349685, -2.591896, -0.770808, 1.570796, 2.110507],accel_mss,speed_ms,0,blend_radius_m)
  movel([0.541557, -1.350126, -2.591603, -0.770660, 1.570796, 2.112353],accel_mss,speed_ms,0,blend_radius_m)
  movel([0.543144, -1.351113, -2.590948, -0.770328, 1.570796, 2.113940],accel_mss,speed_ms,0,blend_radius_m)
  movel([0.544426, -1.352693, -2.589896, -0.769799, 1.570796, 2.115222],accel_mss,speed_ms,0,blend_radius_m)
  movel([0.545344, -1.355662, -2.587911, -0.768816, 1.570796, 2.116140],accel_mss,speed_ms,0,blend_radius_m)
  movel([0.544964, -1.358955, -2.585695, -0.767739, 1.570796, 2.115761],accel_mss,speed_ms,0,blend_radius_m)
  movel([0.543444, -1.362433, -2.583337, -0.766619, 1.570796, 2.114241],accel_mss,speed_ms,0,blend_radius_m)
  movel([0.540946, -1.365969, -2.580923, -0.765497, 1.570796, 2.111742],accel_mss,speed_ms,0,blend_radius_m)
  movel([0.537396, -1.369537, -2.578469, -0.764383, 1.570796, 2.108193],accel_mss,speed_ms,0,blend_radius_m)
  movel([0.533774, -1.371973, -2.576783, -0.763633, 1.570796, 2.104571],accel_mss,speed_ms,0,blend_radius_m)
  movel([0.530140, -1.373419, -2.575779, -0.763191, 1.570796, 2.100936],accel_mss,speed_ms,0,blend_radius_m)
  speed_ms = 0.003
  movel([0.530140, -1.366842, -2.572748, -0.772799, 1.570796, 2.100936],accel_mss,speed_ms,0,blend_radius_m)
  speed_ms = 0.03
  movel([0.530140, -1.341533, -2.560339, -0.810516, 1.570796, 2.100936],accel_mss,speed_ms,0,blend_radius_m)
  #M_RunCode9
  movel([0.640298, -1.231387, -2.625727, -0.855275, 1.570796, 2.211094],accel_mss,speed_ms,0,blend_radius_m)
  #M_RunCode3
  movel([0.640298, -1.258375, -2.639579, -0.814435, 1.570796, 2.211094],accel_mss,speed_ms,0,blend_radius_m)
  speed_ms = 0.003
  movel([0.640298, -1.265443, -2.642973, -0.803973, 1.570796, 2.211094],accel_mss,speed_ms,0,blend_radius_m)
  speed_ms = 0.007
  movel([0.638995, -1.263852, -2.643851, -0.804686, 1.570796, 2.209791],accel_mss,speed_ms,0,blend_radius_m)
  movel([0.638305, -1.261726, -2.645018, -0.805645, 1.570796, 2.209101],accel_mss,speed_ms,0,blend_radius_m)
  movel([0.637965, -1.259330, -2.646327, -0.806732, 1.570796, 2.208761],accel_mss,speed_ms,0,blend_radius_m)
  movel([0.639032, -1.259079, -2.646464, -0.806846, 1.570796, 2.209828],accel_mss,speed_ms,0,blend_radius_m)
  movel([0.639610, -1.259574, -2.646194, -0.806621, 1.570796, 2.210407],accel_mss,speed_ms,0,blend_radius_m)
  movel([0.640340, -1.260082, -2.645917, -0.806390, 1.570796, 2.211136],accel_mss,speed_ms,0,blend_radius_m)
  movel([0.641866, -1.259868, -2.646034, -0.806487, 1.570796, 2.212662],accel_mss,speed_ms,0,blend_radius_m)
  movel([0.643609, -1.258954, -2.646532, -0.806903, 1.570796, 2.214405],accel_mss,speed_ms,0,blend_radius_m)
  movel([0.645309, -1.257727, -2.647199, -0.807463, 1.570796, 2.216105],accel_mss,speed_ms,0,blend_radius_m)
  movel([0.647646, -1.255946, -2.648164, -0.808279, 1.570796, 2.218442],accel_mss,speed_ms,0,blend_radius_m)
  movel([0.647422, -1.252814, -2.649852, -0.809723, 1.570796, 2.218218],accel_mss,speed_ms,0,blend_radius_m)
  movel([0.646332, -1.250712, -2.650978, -0.810699, 1.570796, 2.217128],accel_mss,speed_ms,0,blend_radius_m)
  movel([0.645371, -1.250204, -2.651250, -0.810935, 1.570796, 2.216168],accel_mss,speed_ms,0,blend_radius_m)
  movel([0.644092, -1.250134, -2.651287, -0.810968, 1.570796, 2.214889],accel_mss,speed_ms,0,blend_radius_m)
  movel([0.642462, -1.250567, -2.651056, -0.810766, 1.570796, 2.213258],accel_mss,speed_ms,0,blend_radius_m)
  movel([0.640448, -1.251559, -2.650525, -0.810305, 1.570796, 2.211245],accel_mss,speed_ms,0,blend_radius_m)
  movel([0.641342, -1.249452, -2.651651, -0.811286, 1.570796, 2.212139],accel_mss,speed_ms,0,blend_radius_m)
  movel([0.642348, -1.247651, -2.652609, -0.812129, 1.570796, 2.213144],accel_mss,speed_ms,0,blend_radius_m)
  movel([0.642929, -1.247029, -2.652939, -0.812421, 1.570796, 2.213726],accel_mss,speed_ms,0,blend_radius_m)
  movel([0.643592, -1.246674, -2.653127, -0.812588, 1.570796, 2.214388],accel_mss,speed_ms,0,blend_radius_m)
  movel([0.645206, -1.247042, -2.652932, -0.812415, 1.570796, 2.216003],accel_mss,speed_ms,0,blend_radius_m)
  movel([0.647516, -1.249183, -2.651794, -0.811412, 1.570796, 2.218312],accel_mss,speed_ms,0,blend_radius_m)
  movel([0.649003, -1.252129, -2.650220, -0.810040, 1.570796, 2.219800],accel_mss,speed_ms,0,blend_radius_m)
  movel([0.649248, -1.253833, -2.649304, -0.809252, 1.570796, 2.220044],accel_mss,speed_ms,0,blend_radius_m)
  movel([0.649062, -1.255652, -2.648323, -0.808414, 1.570796, 2.219858],accel_mss,speed_ms,0,blend_radius_m)
  movel([0.648379, -1.257555, -2.647293, -0.807542, 1.570796, 2.219175],accel_mss,speed_ms,0,blend_radius_m)
  movel([0.647119, -1.259514, -2.646227, -0.806648, 1.570796, 2.217916],accel_mss,speed_ms,0,blend_radius_m)
  movel([0.645603, -1.258249, -2.646915, -0.807224, 1.570796, 2.216399],accel_mss,speed_ms,0,blend_radius_m)
  movel([0.642477, -1.266242, -2.642532, -0.803615, 1.570796, 2.213273],accel_mss,speed_ms,0,blend_radius_m)
  movel([0.640298, -1.265443, -2.642973, -0.803973, 1.570796, 2.211094],accel_mss,speed_ms,0,blend_radius_m)
  speed_ms = 0.003
  movel([0.640298, -1.258375, -2.639579, -0.814435, 1.570796, 2.211094],accel_mss,speed_ms,0,blend_radius_m)
  speed_ms = 0.03
  movel([0.640298, -1.231387, -2.625727, -0.855275, 1.570796, 2.211094],accel_mss,speed_ms,0,blend_radius_m)
  #M_RunCode9
  movel([0.618612, -1.173916, -2.654181, -0.884292, 1.570796, 2.189408],accel_mss,speed_ms,0,blend_radius_m)
  #M_RunCode3
  movel([0.618612, -1.201485, -2.668794, -0.842111, 1.570796, 2.189408],accel_mss,speed_ms,0,blend_radius_m)
  speed_ms = 0.003
  movel([0.618612, -1.208739, -2.672382, -0.831268, 1.570796, 2.189408],accel_mss,speed_ms,0,blend_radius_m)
  speed_ms = 0.007
  movel([0.614986, -1.211302, -2.671133, -0.829954, 1.570796, 2.185782],accel_mss,speed_ms,0,blend_radius_m)
  movel([0.611222, -1.213541, -2.670035, -0.828812, 1.570796, 2.182019],accel_mss,speed_ms,0,blend_radius_m)
  movel([0.607365, -1.215415, -2.669113, -0.827861, 1.570796, 2.178161],accel_mss,speed_ms,0,blend_radius_m)
  movel([0.603453, -1.216880, -2.668389, -0.827120, 1.570796, 2.174249],accel_mss,speed_ms,0,blend_radius_m)
  movel([0.599524, -1.217900, -2.667883, -0.826606, 1.570796, 2.170321],accel_mss,speed_ms,0,blend_radius_m)
  movel([0.597567, -1.218004, -2.667832, -0.826554, 1.570796, 2.168364],accel_mss,speed_ms,0,blend_radius_m)
  movel([0.595641, -1.217778, -2.667944, -0.826667, 1.570796, 2.166437],accel_mss,speed_ms,0,blend_radius_m)
  movel([0.593903, -1.217590, -2.668037, -0.826762, 1.570796, 2.164700],accel_mss,speed_ms,0,blend_radius_m)
  movel([0.592520, -1.217799, -2.667933, -0.826657, 1.570796, 2.163316],accel_mss,speed_ms,0,blend_radius_m)
  movel([0.590105, -1.219420, -2.667128, -0.825841, 1.570796, 2.160901],accel_mss,speed_ms,0,blend_radius_m)
  movel([0.586904, -1.222059, -2.665810, -0.824521, 1.570796, 2.157700],accel_mss,speed_ms,0,blend_radius_m)
  movel([0.583585, -1.224846, -2.664409, -0.823134, 1.570796, 2.154381],accel_mss,speed_ms,0,blend_radius_m)
  movel([0.580795, -1.226922, -2.663359, -0.822107, 1.570796, 2.151591],accel_mss,speed_ms,0,blend_radius_m)
  movel([0.575320, -1.229928, -2.661831, -0.820629, 1.570796, 2.146116],accel_mss,speed_ms,0,blend_radius_m)
  movel([0.570456, -1.231825, -2.660862, -0.819702, 1.570796, 2.141252],accel_mss,speed_ms,0,blend_radius_m)
  movel([0.566144, -1.232724, -2.660401, -0.819264, 1.570796, 2.136940],accel_mss,speed_ms,0,blend_radius_m)
  movel([0.562329, -1.232730, -2.660398, -0.819261, 1.570796, 2.133126],accel_mss,speed_ms,0,blend_radius_m)
  movel([0.558962, -1.231946, -2.660800, -0.819643, 1.570796, 2.129758],accel_mss,speed_ms,0,blend_radius_m)
  movel([0.555993, -1.230470, -2.661555, -0.820364, 1.570796, 2.126790],accel_mss,speed_ms,0,blend_radius_m)
  movel([0.553381, -1.228398, -2.662611, -0.821380, 1.570796, 2.124178],accel_mss,speed_ms,0,blend_radius_m)
  movel([0.551085, -1.225828, -2.663913, -0.822648, 1.570796, 2.121881],accel_mss,speed_ms,0,blend_radius_m)
  movel([0.547264, -1.219575, -2.667050, -0.825764, 1.570796, 2.118060],accel_mss,speed_ms,0,blend_radius_m)
  movel([0.544218, -1.212495, -2.670549, -0.829345, 1.570796, 2.115014],accel_mss,speed_ms,0,blend_radius_m)
  movel([0.539198, -1.199145, -2.676993, -0.836251, 1.570796, 2.109994],accel_mss,speed_ms,0,blend_radius_m)
  movel([0.536271, -1.193758, -2.679537, -0.839093, 1.570796, 2.107067],accel_mss,speed_ms,0,blend_radius_m)
  movel([0.532156, -1.188087, -2.682182, -0.842119, 1.570796, 2.102952],accel_mss,speed_ms,0,blend_radius_m)
  movel([0.527012, -1.182480, -2.684763, -0.845146, 1.570796, 2.097808],accel_mss,speed_ms,0,blend_radius_m)
  movel([0.521006, -1.177294, -2.687120, -0.847974, 1.570796, 2.091802],accel_mss,speed_ms,0,blend_radius_m)
  movel([0.514323, -1.172889, -2.689101, -0.850400, 1.570796, 2.085119],accel_mss,speed_ms,0,blend_radius_m)
  movel([0.507165, -1.169614, -2.690559, -0.852216, 1.570796, 2.077962],accel_mss,speed_ms,0,blend_radius_m)
  movel([0.499763, -1.167809, -2.691359, -0.853222, 1.570796, 2.070559],accel_mss,speed_ms,0,blend_radius_m)
  movel([0.496042, -1.167559, -2.691469, -0.853361, 1.570796, 2.066839],accel_mss,speed_ms,0,blend_radius_m)
  movel([0.492354, -1.167794, -2.691365, -0.853230, 1.570796, 2.063150],accel_mss,speed_ms,0,blend_radius_m)
  movel([0.488378, -1.168550, -2.691031, -0.852808, 1.570796, 2.059174],accel_mss,speed_ms,0,blend_radius_m)
  movel([0.483602, -1.169907, -2.690429, -0.852053, 1.570796, 2.054398],accel_mss,speed_ms,0,blend_radius_m)
  movel([0.478305, -1.171902, -2.689542, -0.850946, 1.570796, 2.049102],accel_mss,speed_ms,0,blend_radius_m)
  movel([0.472761, -1.174553, -2.688355, -0.849481, 1.570796, 2.043557],accel_mss,speed_ms,0,blend_radius_m)
  movel([0.467250, -1.177875, -2.686858, -0.847656, 1.570796, 2.038047],accel_mss,speed_ms,0,blend_radius_m)
  movel([0.462053, -1.181881, -2.685037, -0.845471, 1.570796, 2.032850],accel_mss,speed_ms,0,blend_radius_m)
  movel([0.457444, -1.186569, -2.682885, -0.842936, 1.570796, 2.028240],accel_mss,speed_ms,0,blend_radius_m)
  movel([0.455447, -1.189167, -2.681681, -0.841541, 1.570796, 2.026244],accel_mss,speed_ms,0,blend_radius_m)
  movel([0.453700, -1.191937, -2.680391, -0.840061, 1.570796, 2.024496],accel_mss,speed_ms,0,blend_radius_m)
  movel([0.451780, -1.196256, -2.678361, -0.837771, 1.570796, 2.022576],accel_mss,speed_ms,0,blend_radius_m)
  movel([0.451209, -1.199902, -2.676633, -0.835854, 1.570796, 2.022005],accel_mss,speed_ms,0,blend_radius_m)
  movel([0.451821, -1.202946, -2.675179, -0.834265, 1.570796, 2.022618],accel_mss,speed_ms,0,blend_radius_m)
  movel([0.453472, -1.205452, -2.673973, -0.832964, 1.570796, 2.024268],accel_mss,speed_ms,0,blend_radius_m)
  movel([0.456012, -1.207487, -2.672989, -0.831912, 1.570796, 2.026809],accel_mss,speed_ms,0,blend_radius_m)
  movel([0.459296, -1.209115, -2.672199, -0.831075, 1.570796, 2.030092],accel_mss,speed_ms,0,blend_radius_m)
  movel([0.463179, -1.210399, -2.671574, -0.830416, 1.570796, 2.033976],accel_mss,speed_ms,0,blend_radius_m)
  movel([0.467527, -1.211393, -2.671088, -0.829908, 1.570796, 2.038323],accel_mss,speed_ms,0,blend_radius_m)
  movel([0.477053, -1.212735, -2.670431, -0.829223, 1.570796, 2.047849],accel_mss,speed_ms,0,blend_radius_m)
  movel([0.486776, -1.213553, -2.670030, -0.828806, 1.570796, 2.057572],accel_mss,speed_ms,0,blend_radius_m)
  movel([0.495617, -1.214212, -2.669706, -0.828471, 1.570796, 2.066413],accel_mss,speed_ms,0,blend_radius_m)
  movel([0.502493, -1.215038, -2.669299, -0.828052, 1.570796, 2.073289],accel_mss,speed_ms,0,blend_radius_m)
  movel([0.518571, -1.217986, -2.667840, -0.826562, 1.570796, 2.089368],accel_mss,speed_ms,0,blend_radius_m)
  movel([0.526929, -1.219924, -2.666876, -0.825588, 1.570796, 2.097725],accel_mss,speed_ms,0,blend_radius_m)
  movel([0.533101, -1.221975, -2.665852, -0.824563, 1.570796, 2.103897],accel_mss,speed_ms,0,blend_radius_m)
  movel([0.535202, -1.223191, -2.665242, -0.823956, 1.570796, 2.105998],accel_mss,speed_ms,0,blend_radius_m)
  movel([0.536942, -1.224731, -2.664467, -0.823191, 1.570796, 2.107738],accel_mss,speed_ms,0,blend_radius_m)
  movel([0.539386, -1.228658, -2.662479, -0.821253, 1.570796, 2.110183],accel_mss,speed_ms,0,blend_radius_m)
  movel([0.540568, -1.233492, -2.660007, -0.818891, 1.570796, 2.111365],accel_mss,speed_ms,0,blend_radius_m)
  movel([0.540617, -1.238979, -2.657168, -0.816242, 1.570796, 2.111414],accel_mss,speed_ms,0,blend_radius_m)
  movel([0.539672, -1.244871, -2.654080, -0.813438, 1.570796, 2.110468],accel_mss,speed_ms,0,blend_radius_m)
  movel([0.537866, -1.250933, -2.650860, -0.810596, 1.570796, 2.108662],accel_mss,speed_ms,0,blend_radius_m)
  movel([0.535326, -1.256940, -2.647626, -0.807823, 1.570796, 2.106122],accel_mss,speed_ms,0,blend_radius_m)
  movel([0.532174, -1.262673, -2.644499, -0.805217, 1.570796, 2.102971],accel_mss,speed_ms,0,blend_radius_m)
  movel([0.527492, -1.269352, -2.640805, -0.802232, 1.570796, 2.098288],accel_mss,speed_ms,0,blend_radius_m)
  movel([0.525201, -1.271971, -2.639341, -0.801077, 1.570796, 2.095998],accel_mss,speed_ms,0,blend_radius_m)
  movel([0.522923, -1.274178, -2.638101, -0.800109, 1.570796, 2.093719],accel_mss,speed_ms,0,blend_radius_m)
  movel([0.520641, -1.276025, -2.637059, -0.799305, 1.570796, 2.091437],accel_mss,speed_ms,0,blend_radius_m)
  movel([0.518340, -1.277557, -2.636191, -0.798641, 1.570796, 2.089136],accel_mss,speed_ms,0,blend_radius_m)
  movel([0.513623, -1.279858, -2.634883, -0.797649, 1.570796, 2.084419],accel_mss,speed_ms,0,blend_radius_m)
  movel([0.508662, -1.281449, -2.633974, -0.796967, 1.570796, 2.079458],accel_mss,speed_ms,0,blend_radius_m)
  movel([0.503345, -1.282691, -2.633262, -0.796436, 1.570796, 2.074142],accel_mss,speed_ms,0,blend_radius_m)
  movel([0.491275, -1.285528, -2.631629, -0.795232, 1.570796, 2.062071],accel_mss,speed_ms,0,blend_radius_m)
  movel([0.490643, -1.285734, -2.631510, -0.795145, 1.570796, 2.061440],accel_mss,speed_ms,0,blend_radius_m)
  movel([0.490838, -1.285861, -2.631437, -0.795092, 1.570796, 2.061634],accel_mss,speed_ms,0,blend_radius_m)
  movel([0.493262, -1.285926, -2.631399, -0.795064, 1.570796, 2.064059],accel_mss,speed_ms,0,blend_radius_m)
  movel([0.503245, -1.285616, -2.631578, -0.795195, 1.570796, 2.074041],accel_mss,speed_ms,0,blend_radius_m)
  movel([0.519748, -1.285275, -2.631775, -0.795339, 1.570796, 2.090544],accel_mss,speed_ms,0,blend_radius_m)
  movel([0.509882, -1.289690, -2.629214, -0.793484, 1.570796, 2.080678],accel_mss,speed_ms,0,blend_radius_m)
  movel([0.498941, -1.294129, -2.626615, -0.791644, 1.570796, 2.069737],accel_mss,speed_ms,0,blend_radius_m)
  movel([0.487316, -1.298510, -2.624026, -0.789854, 1.570796, 2.058112],accel_mss,speed_ms,0,blend_radius_m)
  movel([0.475394, -1.302746, -2.621498, -0.788145, 1.570796, 2.046190],accel_mss,speed_ms,0,blend_radius_m)
  movel([0.452187, -1.310369, -2.616890, -0.785130, 1.570796, 2.022983],accel_mss,speed_ms,0,blend_radius_m)
  movel([0.441652, -1.313524, -2.614961, -0.783905, 1.570796, 2.012448],accel_mss,speed_ms,0,blend_radius_m)
  movel([0.432328, -1.316069, -2.613395, -0.782925, 1.570796, 2.003124],accel_mss,speed_ms,0,blend_radius_m)
  movel([0.419237, -1.324479, -2.608159, -0.779751, 1.570796, 1.990033],accel_mss,speed_ms,0,blend_radius_m)
  movel([0.406061, -1.333637, -2.602350, -0.776402, 1.570796, 1.976858],accel_mss,speed_ms,0,blend_radius_m)
  movel([0.379896, -1.352852, -2.589790, -0.769746, 1.570796, 1.950693],accel_mss,speed_ms,0,blend_radius_m)
  movel([0.367078, -1.362296, -2.583431, -0.766663, 1.570796, 1.937874],accel_mss,speed_ms,0,blend_radius_m)
  movel([0.354519, -1.371253, -2.577282, -0.763854, 1.570796, 1.925316],accel_mss,speed_ms,0,blend_radius_m)
  movel([0.342251, -1.379465, -2.571545, -0.761378, 1.570796, 1.913048],accel_mss,speed_ms,0,blend_radius_m)
  movel([0.330301, -1.386689, -2.566419, -0.759281, 1.570796, 1.901097],accel_mss,speed_ms,0,blend_radius_m)
  movel([0.325666, -1.389128, -2.564671, -0.758590, 1.570796, 1.896463],accel_mss,speed_ms,0,blend_radius_m)
  movel([0.321263, -1.391100, -2.563252, -0.758037, 1.570796, 1.892059],accel_mss,speed_ms,0,blend_radius_m)
  movel([0.317114, -1.392611, -2.562160, -0.757618, 1.570796, 1.887911],accel_mss,speed_ms,0,blend_radius_m)
  movel([0.313236, -1.393665, -2.561397, -0.757327, 1.570796, 1.884033],accel_mss,speed_ms,0,blend_radius_m)
  movel([0.309656, -1.394263, -2.560963, -0.757163, 1.570796, 1.880452],accel_mss,speed_ms,0,blend_radius_m)
  movel([0.306396, -1.394409, -2.560857, -0.757123, 1.570796, 1.877192],accel_mss,speed_ms,0,blend_radius_m)
  movel([0.303476, -1.394101, -2.561081, -0.757207, 1.570796, 1.874272],accel_mss,speed_ms,0,blend_radius_m)
  movel([0.300924, -1.393343, -2.561630, -0.757416, 1.570796, 1.871720],accel_mss,speed_ms,0,blend_radius_m)
  movel([0.298766, -1.392126, -2.562511, -0.757752, 1.570796, 1.869563],accel_mss,speed_ms,0,blend_radius_m)
  movel([0.297031, -1.390453, -2.563718, -0.758218, 1.570796, 1.867827],accel_mss,speed_ms,0,blend_radius_m)
  movel([0.295743, -1.388318, -2.565252, -0.758818, 1.570796, 1.866539],accel_mss,speed_ms,0,blend_radius_m)
  movel([0.294938, -1.385714, -2.567116, -0.759560, 1.570796, 1.865734],accel_mss,speed_ms,0,blend_radius_m)
  movel([0.294646, -1.382634, -2.569306, -0.760449, 1.570796, 1.865442],accel_mss,speed_ms,0,blend_radius_m)
  movel([0.294902, -1.379073, -2.571821, -0.761494, 1.570796, 1.865699],accel_mss,speed_ms,0,blend_radius_m)
  movel([0.295741, -1.375020, -2.574663, -0.762706, 1.570796, 1.866537],accel_mss,speed_ms,0,blend_radius_m)
  movel([0.297202, -1.370466, -2.577827, -0.764096, 1.570796, 1.867998],accel_mss,speed_ms,0,blend_radius_m)
  movel([0.300876, -1.371718, -2.576960, -0.763711, 1.570796, 1.871673],accel_mss,speed_ms,0,blend_radius_m)
  movel([0.302745, -1.372211, -2.576618, -0.763560, 1.570796, 1.873541],accel_mss,speed_ms,0,blend_radius_m)
  movel([0.304799, -1.372208, -2.576620, -0.763561, 1.570796, 1.875595],accel_mss,speed_ms,0,blend_radius_m)
  movel([0.306575, -1.371659, -2.577001, -0.763729, 1.570796, 1.877371],accel_mss,speed_ms,0,blend_radius_m)
  movel([0.308779, -1.370564, -2.577759, -0.764066, 1.570796, 1.879576],accel_mss,speed_ms,0,blend_radius_m)
  movel([0.314252, -1.366988, -2.580224, -0.765177, 1.570796, 1.885048],accel_mss,speed_ms,0,blend_radius_m)
  movel([0.320765, -1.362012, -2.583623, -0.766754, 1.570796, 1.891561],accel_mss,speed_ms,0,blend_radius_m)
  movel([0.327864, -1.356167, -2.587572, -0.768650, 1.570796, 1.898660],accel_mss,speed_ms,0,blend_radius_m)
  movel([0.341870, -1.344056, -2.595603, -0.772730, 1.570796, 1.912667],accel_mss,speed_ms,0,blend_radius_m)
  movel([0.352135, -1.335193, -2.601352, -0.775844, 1.570796, 1.922931],accel_mss,speed_ms,0,blend_radius_m)
  movel([0.361407, -1.328046, -2.605910, -0.778433, 1.570796, 1.932203],accel_mss,speed_ms,0,blend_radius_m)
  movel([0.370798, -1.320857, -2.610426, -0.781107, 1.570796, 1.941595],accel_mss,speed_ms,0,blend_radius_m)
  movel([0.351774, -1.324841, -2.607932, -0.779616, 1.570796, 1.922571],accel_mss,speed_ms,0,blend_radius_m)
  movel([0.341960, -1.326553, -2.606853, -0.778982, 1.570796, 1.912756],accel_mss,speed_ms,0,blend_radius_m)
  movel([0.332625, -1.327411, -2.606312, -0.778666, 1.570796, 1.903421],accel_mss,speed_ms,0,blend_radius_m)
  movel([0.328292, -1.327360, -2.606344, -0.778685, 1.570796, 1.899088],accel_mss,speed_ms,0,blend_radius_m)
  movel([0.324266, -1.326901, -2.606634, -0.778854, 1.570796, 1.895062],accel_mss,speed_ms,0,blend_radius_m)
  movel([0.320604, -1.325968, -2.607222, -0.779199, 1.570796, 1.891400],accel_mss,speed_ms,0,blend_radius_m)
  movel([0.317373, -1.324491, -2.608152, -0.779747, 1.570796, 1.888169],accel_mss,speed_ms,0,blend_radius_m)
  movel([0.314634, -1.322395, -2.609465, -0.780529, 1.570796, 1.885430],accel_mss,speed_ms,0,blend_radius_m)
  movel([0.312446, -1.319613, -2.611200, -0.781576, 1.570796, 1.883243],accel_mss,speed_ms,0,blend_radius_m)
  movel([0.310885, -1.316063, -2.613399, -0.782928, 1.570796, 1.881681],accel_mss,speed_ms,0,blend_radius_m)
  movel([0.310014, -1.311659, -2.616102, -0.784627, 1.570796, 1.880810],accel_mss,speed_ms,0,blend_radius_m)
  movel([0.310106, -1.305931, -2.619582, -0.786876, 1.570796, 1.880903],accel_mss,speed_ms,0,blend_radius_m)
  movel([0.311426, -1.299633, -2.623357, -0.789398, 1.570796, 1.882222],accel_mss,speed_ms,0,blend_radius_m)
  movel([0.313888, -1.292959, -2.627303, -0.792127, 1.570796, 1.884684],accel_mss,speed_ms,0,blend_radius_m)
  movel([0.317395, -1.286115, -2.631290, -0.794984, 1.570796, 1.888191],accel_mss,speed_ms,0,blend_radius_m)
  movel([0.321852, -1.279319, -2.635189, -0.797880, 1.570796, 1.892648],accel_mss,speed_ms,0,blend_radius_m)
  movel([0.327144, -1.272806, -2.638873, -0.800710, 1.570796, 1.897940],accel_mss,speed_ms,0,blend_radius_m)
  movel([0.333157, -1.266816, -2.642214, -0.803359, 1.570796, 1.903953],accel_mss,speed_ms,0,blend_radius_m)
  movel([0.339761, -1.261607, -2.645083, -0.805699, 1.570796, 1.910557],accel_mss,speed_ms,0,blend_radius_m)
  movel([0.343560, -1.259552, -2.646206, -0.806631, 1.570796, 1.914356],accel_mss,speed_ms,0,blend_radius_m)
  movel([0.347804, -1.258080, -2.647007, -0.807302, 1.570796, 1.918601],accel_mss,speed_ms,0,blend_radius_m)
  movel([0.351133, -1.257735, -2.647195, -0.807459, 1.570796, 1.921929],accel_mss,speed_ms,0,blend_radius_m)
  movel([0.352023, -1.258156, -2.646966, -0.807267, 1.570796, 1.922819],accel_mss,speed_ms,0,blend_radius_m)
  movel([0.352174, -1.259056, -2.646477, -0.806857, 1.570796, 1.922970],accel_mss,speed_ms,0,blend_radius_m)
  movel([0.348824, -1.260160, -2.645875, -0.806355, 1.570796, 1.919620],accel_mss,speed_ms,0,blend_radius_m)
  movel([0.345957, -1.261443, -2.645173, -0.805773, 1.570796, 1.916754],accel_mss,speed_ms,0,blend_radius_m)
  movel([0.343566, -1.262869, -2.644391, -0.805129, 1.570796, 1.914362],accel_mss,speed_ms,0,blend_radius_m)
  movel([0.341628, -1.264406, -2.643546, -0.804437, 1.570796, 1.912424],accel_mss,speed_ms,0,blend_radius_m)
  movel([0.340128, -1.266024, -2.642652, -0.803713, 1.570796, 1.910924],accel_mss,speed_ms,0,blend_radius_m)
  movel([0.339052, -1.267689, -2.641729, -0.802970, 1.570796, 1.909848],accel_mss,speed_ms,0,blend_radius_m)
  movel([0.338377, -1.269375, -2.640792, -0.802222, 1.570796, 1.909173],accel_mss,speed_ms,0,blend_radius_m)
  movel([0.338090, -1.271052, -2.639856, -0.801481, 1.570796, 1.908887],accel_mss,speed_ms,0,blend_radius_m)
  movel([0.338601, -1.274269, -2.638050, -0.800070, 1.570796, 1.909397],accel_mss,speed_ms,0,blend_radius_m)
  movel([0.340435, -1.277118, -2.636440, -0.798831, 1.570796, 1.911232],accel_mss,speed_ms,0,blend_radius_m)
  movel([0.343451, -1.279397, -2.635145, -0.797847, 1.570796, 1.914248],accel_mss,speed_ms,0,blend_radius_m)
  movel([0.347518, -1.280888, -2.634295, -0.797207, 1.570796, 1.918315],accel_mss,speed_ms,0,blend_radius_m)
  movel([0.350339, -1.281223, -2.634103, -0.797063, 1.570796, 1.921136],accel_mss,speed_ms,0,blend_radius_m)
  movel([0.353952, -1.281188, -2.634123, -0.797078, 1.570796, 1.924749],accel_mss,speed_ms,0,blend_radius_m)
  movel([0.363138, -1.280187, -2.634695, -0.797507, 1.570796, 1.933935],accel_mss,speed_ms,0,blend_radius_m)
  movel([0.374236, -1.278244, -2.635801, -0.798344, 1.570796, 1.945033],accel_mss,speed_ms,0,blend_radius_m)
  movel([0.386417, -1.275704, -2.637241, -0.799445, 1.570796, 1.957214],accel_mss,speed_ms,0,blend_radius_m)
  movel([0.410657, -1.270074, -2.640402, -0.801913, 1.570796, 1.981453],accel_mss,speed_ms,0,blend_radius_m)
  movel([0.429065, -1.265519, -2.642931, -0.803938, 1.570796, 1.999862],accel_mss,speed_ms,0,blend_radius_m)
  movel([0.438346, -1.263231, -2.644192, -0.804966, 1.570796, 2.009142],accel_mss,speed_ms,0,blend_radius_m)
  movel([0.443381, -1.261840, -2.644956, -0.805594, 1.570796, 2.014178],accel_mss,speed_ms,0,blend_radius_m)
  movel([0.447252, -1.260440, -2.645721, -0.806227, 1.570796, 2.018048],accel_mss,speed_ms,0,blend_radius_m)
  movel([0.448324, -1.259833, -2.646053, -0.806503, 1.570796, 2.019120],accel_mss,speed_ms,0,blend_radius_m)
  movel([0.448774, -1.259284, -2.646352, -0.806753, 1.570796, 2.019571],accel_mss,speed_ms,0,blend_radius_m)
  movel([0.448312, -1.258068, -2.647014, -0.807307, 1.570796, 2.019108],accel_mss,speed_ms,0,blend_radius_m)
  movel([0.445522, -1.255611, -2.648345, -0.808433, 1.570796, 2.016318],accel_mss,speed_ms,0,blend_radius_m)
  movel([0.441913, -1.253827, -2.649308, -0.809255, 1.570796, 2.012709],accel_mss,speed_ms,0,blend_radius_m)
  movel([0.433762, -1.250480, -2.651102, -0.810807, 1.570796, 2.004558],accel_mss,speed_ms,0,blend_radius_m)
  movel([0.429980, -1.247995, -2.652426, -0.811968, 1.570796, 2.000776],accel_mss,speed_ms,0,blend_radius_m)
  movel([0.426898, -1.244335, -2.654363, -0.813692, 1.570796, 1.997694],accel_mss,speed_ms,0,blend_radius_m)
  movel([0.425739, -1.241911, -2.655636, -0.814842, 1.570796, 1.996536],accel_mss,speed_ms,0,blend_radius_m)
  movel([0.424901, -1.238999, -2.657157, -0.816232, 1.570796, 1.995697],accel_mss,speed_ms,0,blend_radius_m)
  movel([0.424432, -1.235539, -2.658951, -0.817898, 1.570796, 1.995229],accel_mss,speed_ms,0,blend_radius_m)
  movel([0.424388, -1.231460, -2.661049, -0.819880, 1.570796, 1.995185],accel_mss,speed_ms,0,blend_radius_m)
  movel([0.425174, -1.225716, -2.663970, -0.822703, 1.570796, 1.995970],accel_mss,speed_ms,0,blend_radius_m)
  movel([0.426979, -1.219930, -2.666874, -0.825586, 1.570796, 1.997775],accel_mss,speed_ms,0,blend_radius_m)
  movel([0.429691, -1.214126, -2.669748, -0.828515, 1.570796, 2.000487],accel_mss,speed_ms,0,blend_radius_m)
  movel([0.433204, -1.208325, -2.672583, -0.831481, 1.570796, 2.004001],accel_mss,speed_ms,0,blend_radius_m)
  movel([0.437393, -1.202554, -2.675366, -0.834469, 1.570796, 2.008189],accel_mss,speed_ms,0,blend_radius_m)
  movel([0.442138, -1.196845, -2.678083, -0.837461, 1.570796, 2.012934],accel_mss,speed_ms,0,blend_radius_m)
  movel([0.447315, -1.191224, -2.680724, -0.840441, 1.570796, 2.018111],accel_mss,speed_ms,0,blend_radius_m)
  movel([0.452799, -1.185726, -2.683273, -0.843390, 1.570796, 2.023596],accel_mss,speed_ms,0,blend_radius_m)
  movel([0.463644, -1.175989, -2.687709, -0.848691, 1.570796, 2.034440],accel_mss,speed_ms,0,blend_radius_m)
  movel([0.473616, -1.168330, -2.691128, -0.852931, 1.570796, 2.044412],accel_mss,speed_ms,0,blend_radius_m)
  movel([0.482210, -1.162670, -2.693616, -0.856103, 1.570796, 2.053006],accel_mss,speed_ms,0,blend_radius_m)
  movel([0.488934, -1.158899, -2.695255, -0.858235, 1.570796, 2.059730],accel_mss,speed_ms,0,blend_radius_m)
  movel([0.498877, -1.154497, -2.697150, -0.860743, 1.570796, 2.069673],accel_mss,speed_ms,0,blend_radius_m)
  movel([0.508411, -1.151584, -2.698393, -0.862412, 1.570796, 2.079207],accel_mss,speed_ms,0,blend_radius_m)
  movel([0.517405, -1.150134, -2.699008, -0.863247, 1.570796, 2.088201],accel_mss,speed_ms,0,blend_radius_m)
  movel([0.525733, -1.150119, -2.699015, -0.863255, 1.570796, 2.096529],accel_mss,speed_ms,0,blend_radius_m)
  movel([0.533278, -1.151486, -2.698434, -0.862468, 1.570796, 2.104075],accel_mss,speed_ms,0,blend_radius_m)
  movel([0.539930, -1.154176, -2.697287, -0.860926, 1.570796, 2.110726],accel_mss,speed_ms,0,blend_radius_m)
  movel([0.545599, -1.158106, -2.695598, -0.858686, 1.570796, 2.116396],accel_mss,speed_ms,0,blend_radius_m)
  movel([0.550201, -1.163189, -2.693389, -0.855811, 1.570796, 2.120997],accel_mss,speed_ms,0,blend_radius_m)
  movel([0.553359, -1.168678, -2.690974, -0.852737, 1.570796, 2.124156],accel_mss,speed_ms,0,blend_radius_m)
  movel([0.555869, -1.174627, -2.688322, -0.849440, 1.570796, 2.126665],accel_mss,speed_ms,0,blend_radius_m)
  movel([0.558209, -1.180541, -2.685648, -0.846200, 1.570796, 2.129005],accel_mss,speed_ms,0,blend_radius_m)
  movel([0.560863, -1.185964, -2.683164, -0.843262, 1.570796, 2.131659],accel_mss,speed_ms,0,blend_radius_m)
  movel([0.564292, -1.190448, -2.681086, -0.840856, 1.570796, 2.135088],accel_mss,speed_ms,0,blend_radius_m)
  movel([0.566444, -1.192205, -2.680265, -0.839919, 1.570796, 2.137241],accel_mss,speed_ms,0,blend_radius_m)
  movel([0.568968, -1.193569, -2.679626, -0.839194, 1.570796, 2.139764],accel_mss,speed_ms,0,blend_radius_m)
  movel([0.571917, -1.194490, -2.679194, -0.838706, 1.570796, 2.142713],accel_mss,speed_ms,0,blend_radius_m)
  movel([0.575354, -1.194916, -2.678993, -0.838480, 1.570796, 2.146150],accel_mss,speed_ms,0,blend_radius_m)
  movel([0.579344, -1.194790, -2.679052, -0.838546, 1.570796, 2.150140],accel_mss,speed_ms,0,blend_radius_m)
  movel([0.583943, -1.194069, -2.679392, -0.838929, 1.570796, 2.154740],accel_mss,speed_ms,0,blend_radius_m)
  movel([0.588161, -1.192792, -2.679991, -0.839606, 1.570796, 2.158957],accel_mss,speed_ms,0,blend_radius_m)
  movel([0.591903, -1.190918, -2.680866, -0.840604, 1.570796, 2.162699],accel_mss,speed_ms,0,blend_radius_m)
  movel([0.595162, -1.188555, -2.681965, -0.841869, 1.570796, 2.165958],accel_mss,speed_ms,0,blend_radius_m)
  movel([0.597932, -1.185817, -2.683231, -0.843341, 1.570796, 2.168728],accel_mss,speed_ms,0,blend_radius_m)
  movel([0.600197, -1.182817, -2.684609, -0.844963, 1.570796, 2.170993],accel_mss,speed_ms,0,blend_radius_m)
  movel([0.601941, -1.179676, -2.686041, -0.846671, 1.570796, 2.172737],accel_mss,speed_ms,0,blend_radius_m)
  movel([0.603151, -1.176514, -2.687473, -0.848403, 1.570796, 2.173948],accel_mss,speed_ms,0,blend_radius_m)
  movel([0.603802, -1.173459, -2.688845, -0.850084, 1.570796, 2.174598],accel_mss,speed_ms,0,blend_radius_m)
  movel([0.603875, -1.170638, -2.690104, -0.851646, 1.570796, 2.174671],accel_mss,speed_ms,0,blend_radius_m)
  movel([0.603353, -1.168186, -2.691192, -0.853011, 1.570796, 2.174149],accel_mss,speed_ms,0,blend_radius_m)
  movel([0.602213, -1.166236, -2.692052, -0.854100, 1.570796, 2.173010],accel_mss,speed_ms,0,blend_radius_m)
  movel([0.600441, -1.164921, -2.692630, -0.854838, 1.570796, 2.171238],accel_mss,speed_ms,0,blend_radius_m)
  movel([0.598020, -1.164375, -2.692870, -0.855144, 1.570796, 2.168816],accel_mss,speed_ms,0,blend_radius_m)
  movel([0.594936, -1.164733, -2.692713, -0.854943, 1.570796, 2.165732],accel_mss,speed_ms,0,blend_radius_m)
  movel([0.591188, -1.166116, -2.692105, -0.854168, 1.570796, 2.161985],accel_mss,speed_ms,0,blend_radius_m)
  movel([0.586773, -1.168651, -2.690986, -0.852752, 1.570796, 2.157569],accel_mss,speed_ms,0,blend_radius_m)
  movel([0.589051, -1.169187, -2.690749, -0.852453, 1.570796, 2.159848],accel_mss,speed_ms,0,blend_radius_m)
  movel([0.590621, -1.170198, -2.690300, -0.851891, 1.570796, 2.161418],accel_mss,speed_ms,0,blend_radius_m)
  movel([0.591475, -1.171600, -2.689676, -0.851113, 1.570796, 2.162272],accel_mss,speed_ms,0,blend_radius_m)
  movel([0.591610, -1.173321, -2.688907, -0.850161, 1.570796, 2.162407],accel_mss,speed_ms,0,blend_radius_m)
  movel([0.591022, -1.175290, -2.688024, -0.849075, 1.570796, 2.161818],accel_mss,speed_ms,0,blend_radius_m)
  movel([0.589710, -1.177428, -2.687060, -0.847901, 1.570796, 2.160506],accel_mss,speed_ms,0,blend_radius_m)
  movel([0.587671, -1.179671, -2.686044, -0.846675, 1.570796, 2.158468],accel_mss,speed_ms,0,blend_radius_m)
  movel([0.584904, -1.181948, -2.685006, -0.845435, 1.570796, 2.155700],accel_mss,speed_ms,0,blend_radius_m)
  movel([0.579895, -1.184989, -2.683612, -0.843787, 1.570796, 2.150692],accel_mss,speed_ms,0,blend_radius_m)
  movel([0.575418, -1.186579, -2.682880, -0.842930, 1.570796, 2.146214],accel_mss,speed_ms,0,blend_radius_m)
  movel([0.571478, -1.186871, -2.682745, -0.842773, 1.570796, 2.142275],accel_mss,speed_ms,0,blend_radius_m)
  movel([0.568102, -1.186012, -2.683141, -0.843235, 1.570796, 2.138898],accel_mss,speed_ms,0,blend_radius_m)
  movel([0.565315, -1.184127, -2.684009, -0.844253, 1.570796, 2.136112],accel_mss,speed_ms,0,blend_radius_m)
  movel([0.563152, -1.181348, -2.685280, -0.845761, 1.570796, 2.133948],accel_mss,speed_ms,0,blend_radius_m)
  movel([0.561649, -1.177798, -2.686893, -0.847698, 1.570796, 2.132446],accel_mss,speed_ms,0,blend_radius_m)
  movel([0.560852, -1.173598, -2.688783, -0.850008, 1.570796, 2.131648],accel_mss,speed_ms,0,blend_radius_m)
  movel([0.560803, -1.168872, -2.690888, -0.852629, 1.570796, 2.131600],accel_mss,speed_ms,0,blend_radius_m)
  movel([0.561561, -1.163744, -2.693146, -0.855499, 1.570796, 2.132357],accel_mss,speed_ms,0,blend_radius_m)
  movel([0.563168, -1.158342, -2.695496, -0.858552, 1.570796, 2.133965],accel_mss,speed_ms,0,blend_radius_m)
  movel([0.565684, -1.152800, -2.697875, -0.861714, 1.570796, 2.136480],accel_mss,speed_ms,0,blend_radius_m)
  movel([0.569154, -1.147259, -2.700223, -0.864907, 1.570796, 2.139950],accel_mss,speed_ms,0,blend_radius_m)
  movel([0.573631, -1.141867, -2.702478, -0.868044, 1.570796, 2.144428],accel_mss,speed_ms,0,blend_radius_m)
  movel([0.579156, -1.136786, -2.704577, -0.871026, 1.570796, 2.149952],accel_mss,speed_ms,0,blend_radius_m)
  movel([0.585766, -1.132190, -2.706454, -0.873745, 1.570796, 2.156563],accel_mss,speed_ms,0,blend_radius_m)
  movel([0.590668, -1.129467, -2.707556, -0.875366, 1.570796, 2.161464],accel_mss,speed_ms,0,blend_radius_m)
  movel([0.595527, -1.127201, -2.708468, -0.876720, 1.570796, 2.166323],accel_mss,speed_ms,0,blend_radius_m)
  movel([0.600297, -1.125399, -2.709189, -0.877800, 1.570796, 2.171093],accel_mss,speed_ms,0,blend_radius_m)
  movel([0.604941, -1.124070, -2.709720, -0.878599, 1.570796, 2.175737],accel_mss,speed_ms,0,blend_radius_m)
  movel([0.609409, -1.123228, -2.710055, -0.879106, 1.570796, 2.180205],accel_mss,speed_ms,0,blend_radius_m)
  movel([0.613661, -1.122876, -2.710195, -0.879318, 1.570796, 2.184457],accel_mss,speed_ms,0,blend_radius_m)
  movel([0.617658, -1.123019, -2.710138, -0.879232, 1.570796, 2.188454],accel_mss,speed_ms,0,blend_radius_m)
  movel([0.621360, -1.123657, -2.709884, -0.878848, 1.570796, 2.192156],accel_mss,speed_ms,0,blend_radius_m)
  movel([0.624719, -1.124796, -2.709430, -0.878162, 1.570796, 2.195516],accel_mss,speed_ms,0,blend_radius_m)
  movel([0.627708, -1.126434, -2.708775, -0.877179, 1.570796, 2.198504],accel_mss,speed_ms,0,blend_radius_m)
  movel([0.630282, -1.128567, -2.707919, -0.875903, 1.570796, 2.201078],accel_mss,speed_ms,0,blend_radius_m)
  movel([0.632408, -1.131189, -2.706860, -0.874340, 1.570796, 2.203204],accel_mss,speed_ms,0,blend_radius_m)
  movel([0.634059, -1.134293, -2.705598, -0.872498, 1.570796, 2.204856],accel_mss,speed_ms,0,blend_radius_m)
  movel([0.635195, -1.137877, -2.704129, -0.870384, 1.570796, 2.205991],accel_mss,speed_ms,0,blend_radius_m)
  movel([0.635790, -1.141928, -2.702453, -0.868008, 1.570796, 2.206587],accel_mss,speed_ms,0,blend_radius_m)
  movel([0.635819, -1.146433, -2.700570, -0.865386, 1.570796, 2.206615],accel_mss,speed_ms,0,blend_radius_m)
  movel([0.634733, -1.151374, -2.698482, -0.862533, 1.570796, 2.205529],accel_mss,speed_ms,0,blend_radius_m)
  movel([0.632656, -1.156964, -2.696090, -0.859335, 1.570796, 2.203452],accel_mss,speed_ms,0,blend_radius_m)
  movel([0.630642, -1.161793, -2.693998, -0.856598, 1.570796, 2.201438],accel_mss,speed_ms,0,blend_radius_m)
  movel([0.629715, -1.164497, -2.692816, -0.855075, 1.570796, 2.200511],accel_mss,speed_ms,0,blend_radius_m)
  movel([0.630575, -1.165883, -2.692208, -0.854298, 1.570796, 2.201372],accel_mss,speed_ms,0,blend_radius_m)
  movel([0.632609, -1.167559, -2.691469, -0.853361, 1.570796, 2.203405],accel_mss,speed_ms,0,blend_radius_m)
  movel([0.634843, -1.169409, -2.690650, -0.852330, 1.570796, 2.205639],accel_mss,speed_ms,0,blend_radius_m)
  movel([0.636333, -1.171292, -2.689813, -0.851283, 1.570796, 2.207130],accel_mss,speed_ms,0,blend_radius_m)
  movel([0.637324, -1.174538, -2.688362, -0.849489, 1.570796, 2.208121],accel_mss,speed_ms,0,blend_radius_m)
  movel([0.637636, -1.177970, -2.686815, -0.847604, 1.570796, 2.208432],accel_mss,speed_ms,0,blend_radius_m)
  movel([0.637319, -1.181532, -2.685196, -0.845661, 1.570796, 2.208115],accel_mss,speed_ms,0,blend_radius_m)
  movel([0.636436, -1.185170, -2.683529, -0.843690, 1.570796, 2.207232],accel_mss,speed_ms,0,blend_radius_m)
  movel([0.635031, -1.188837, -2.681835, -0.841718, 1.570796, 2.205828],accel_mss,speed_ms,0,blend_radius_m)
  movel([0.633164, -1.192478, -2.680138, -0.839773, 1.570796, 2.203961],accel_mss,speed_ms,0,blend_radius_m)
  movel([0.630887, -1.196048, -2.678460, -0.837881, 1.570796, 2.201683],accel_mss,speed_ms,0,blend_radius_m)
  movel([0.628243, -1.199502, -2.676823, -0.836064, 1.570796, 2.199039],accel_mss,speed_ms,0,blend_radius_m)
  movel([0.625284, -1.202799, -2.675249, -0.834341, 1.570796, 2.196080],accel_mss,speed_ms,0,blend_radius_m)
  movel([0.622061, -1.205890, -2.673762, -0.832737, 1.570796, 2.192857],accel_mss,speed_ms,0,blend_radius_m)
  movel([0.618612, -1.208739, -2.672382, -0.831268, 1.570796, 2.189408],accel_mss,speed_ms,0,blend_radius_m)
  speed_ms = 0.003
  movel([0.618612, -1.201485, -2.668794, -0.842111, 1.570796, 2.189408],accel_mss,speed_ms,0,blend_radius_m)
  speed_ms = 0.03
  movel([0.618612, -1.173916, -2.654181, -0.884292, 1.570796, 2.189408],accel_mss,speed_ms,0,blend_radius_m)
  #M_RunCode9
  movel([0.640733, -1.173424, -2.654409, -0.884556, 1.570796, 2.211529],accel_mss,speed_ms,0,blend_radius_m)
  #M_RunCode3
  movel([0.640733, -1.200996, -2.669029, -0.842364, 1.570796, 2.211529],accel_mss,speed_ms,0,blend_radius_m)
  speed_ms = 0.003
  movel([0.640733, -1.208251, -2.672619, -0.831519, 1.570796, 2.211529],accel_mss,speed_ms,0,blend_radius_m)
  speed_ms = 0.007
  movel([0.642244, -1.205238, -2.674076, -0.833075, 1.570796, 2.213041],accel_mss,speed_ms,0,blend_radius_m)
  movel([0.646083, -1.199130, -2.677000, -0.836259, 1.570796, 2.216879],accel_mss,speed_ms,0,blend_radius_m)
  movel([0.649594, -1.193117, -2.679838, -0.839434, 1.570796, 2.220390],accel_mss,speed_ms,0,blend_radius_m)
  movel([0.650683, -1.190223, -2.681190, -0.840976, 1.570796, 2.221479],accel_mss,speed_ms,0,blend_radius_m)
  movel([0.651033, -1.187450, -2.682477, -0.842462, 1.570796, 2.221829],accel_mss,speed_ms,0,blend_radius_m)
  movel([0.651466, -1.189153, -2.681688, -0.841548, 1.570796, 2.222262],accel_mss,speed_ms,0,blend_radius_m)
  movel([0.651508, -1.192622, -2.680070, -0.839697, 1.570796, 2.222304],accel_mss,speed_ms,0,blend_radius_m)
  movel([0.650665, -1.196121, -2.678425, -0.837843, 1.570796, 2.221462],accel_mss,speed_ms,0,blend_radius_m)
  movel([0.649218, -1.199641, -2.676757, -0.835991, 1.570796, 2.220014],accel_mss,speed_ms,0,blend_radius_m)
  movel([0.647442, -1.203171, -2.675071, -0.834148, 1.570796, 2.218238],accel_mss,speed_ms,0,blend_radius_m)
  movel([0.643977, -1.210227, -2.671658, -0.830504, 1.570796, 2.214773],accel_mss,speed_ms,0,blend_radius_m)
  movel([0.642819, -1.213737, -2.669939, -0.828713, 1.570796, 2.213615],accel_mss,speed_ms,0,blend_radius_m)
  movel([0.642393, -1.217224, -2.668219, -0.826947, 1.570796, 2.213189],accel_mss,speed_ms,0,blend_radius_m)
  movel([0.642722, -1.220825, -2.666427, -0.825137, 1.570796, 2.213518],accel_mss,speed_ms,0,blend_radius_m)
  movel([0.643100, -1.222640, -2.665518, -0.824231, 1.570796, 2.213896],accel_mss,speed_ms,0,blend_radius_m)
  movel([0.643606, -1.223512, -2.665080, -0.823797, 1.570796, 2.214403],accel_mss,speed_ms,0,blend_radius_m)
  movel([0.645568, -1.222876, -2.665400, -0.824113, 1.570796, 2.216364],accel_mss,speed_ms,0,blend_radius_m)
  movel([0.647164, -1.222435, -2.665621, -0.824333, 1.570796, 2.217961],accel_mss,speed_ms,0,blend_radius_m)
  movel([0.648712, -1.222309, -2.665684, -0.824396, 1.570796, 2.219509],accel_mss,speed_ms,0,blend_radius_m)
  movel([0.651419, -1.222824, -2.665426, -0.824139, 1.570796, 2.222216],accel_mss,speed_ms,0,blend_radius_m)
  movel([0.653147, -1.223713, -2.664979, -0.823697, 1.570796, 2.223943],accel_mss,speed_ms,0,blend_radius_m)
  movel([0.654106, -1.224930, -2.664367, -0.823093, 1.570796, 2.224902],accel_mss,speed_ms,0,blend_radius_m)
  movel([0.654502, -1.226430, -2.663609, -0.822351, 1.570796, 2.225299],accel_mss,speed_ms,0,blend_radius_m)
  movel([0.654448, -1.230102, -2.661743, -0.820544, 1.570796, 2.225245],accel_mss,speed_ms,0,blend_radius_m)
  movel([0.654631, -1.234389, -2.659545, -0.818455, 1.570796, 2.225428],accel_mss,speed_ms,0,blend_radius_m)
  movel([0.655939, -1.239593, -2.656848, -0.815948, 1.570796, 2.226735],accel_mss,speed_ms,0,blend_radius_m)
  movel([0.657464, -1.244611, -2.654217, -0.813561, 1.570796, 2.228260],accel_mss,speed_ms,0,blend_radius_m)
  movel([0.658682, -1.249764, -2.651485, -0.811141, 1.570796, 2.229478],accel_mss,speed_ms,0,blend_radius_m)
  movel([0.659082, -1.255356, -2.648483, -0.808550, 1.570796, 2.229878],accel_mss,speed_ms,0,blend_radius_m)
  movel([0.658762, -1.258600, -2.646725, -0.807064, 1.570796, 2.229558],accel_mss,speed_ms,0,blend_radius_m)
  movel([0.658062, -1.261937, -2.644903, -0.805550, 1.570796, 2.228859],accel_mss,speed_ms,0,blend_radius_m)
  movel([0.655919, -1.268743, -2.641144, -0.802502, 1.570796, 2.226716],accel_mss,speed_ms,0,blend_radius_m)
  movel([0.653429, -1.275481, -2.637366, -0.799541, 1.570796, 2.224225],accel_mss,speed_ms,0,blend_radius_m)
  movel([0.651348, -1.281868, -2.633733, -0.796787, 1.570796, 2.222144],accel_mss,speed_ms,0,blend_radius_m)
  movel([0.649216, -1.292077, -2.627820, -0.792492, 1.570796, 2.220013],accel_mss,speed_ms,0,blend_radius_m)
  movel([0.648432, -1.296382, -2.625287, -0.790721, 1.570796, 2.219228],accel_mss,speed_ms,0,blend_radius_m)
  movel([0.647423, -1.300483, -2.622851, -0.789055, 1.570796, 2.218219],accel_mss,speed_ms,0,blend_radius_m)
  movel([0.645886, -1.304624, -2.620369, -0.787395, 1.570796, 2.216682],accel_mss,speed_ms,0,blend_radius_m)
  movel([0.643527, -1.309032, -2.617703, -0.785653, 1.570796, 2.214323],accel_mss,speed_ms,0,blend_radius_m)
  movel([0.640056, -1.313941, -2.614705, -0.783743, 1.570796, 2.210852],accel_mss,speed_ms,0,blend_radius_m)
  movel([0.635201, -1.319570, -2.611227, -0.781593, 1.570796, 2.205997],accel_mss,speed_ms,0,blend_radius_m)
  movel([0.630905, -1.323885, -2.608532, -0.779972, 1.570796, 2.201701],accel_mss,speed_ms,0,blend_radius_m)
  movel([0.626672, -1.327560, -2.606217, -0.778611, 1.570796, 2.197468],accel_mss,speed_ms,0,blend_radius_m)
  movel([0.622498, -1.330640, -2.604264, -0.777485, 1.570796, 2.193294],accel_mss,speed_ms,0,blend_radius_m)
  movel([0.618384, -1.333162, -2.602654, -0.776573, 1.570796, 2.189180],accel_mss,speed_ms,0,blend_radius_m)
  movel([0.614328, -1.335166, -2.601369, -0.775854, 1.570796, 2.185124],accel_mss,speed_ms,0,blend_radius_m)
  movel([0.610329, -1.336687, -2.600390, -0.775312, 1.570796, 2.181125],accel_mss,speed_ms,0,blend_radius_m)
  movel([0.606388, -1.337762, -2.599696, -0.774930, 1.570796, 2.177185],accel_mss,speed_ms,0,blend_radius_m)
  movel([0.602512, -1.338421, -2.599270, -0.774697, 1.570796, 2.173308],accel_mss,speed_ms,0,blend_radius_m)
  movel([0.598700, -1.338696, -2.599092, -0.774601, 1.570796, 2.169497],accel_mss,speed_ms,0,blend_radius_m)
  movel([0.594954, -1.338620, -2.599142, -0.774627, 1.570796, 2.165750],accel_mss,speed_ms,0,blend_radius_m)
  movel([0.587680, -1.337529, -2.599847, -0.775013, 1.570796, 2.158477],accel_mss,speed_ms,0,blend_radius_m)
  movel([0.580737, -1.335374, -2.601235, -0.775779, 1.570796, 2.151534],accel_mss,speed_ms,0,blend_radius_m)
  movel([0.574175, -1.332382, -2.603153, -0.776854, 1.570796, 2.144971],accel_mss,speed_ms,0,blend_radius_m)
  movel([0.568506, -1.328893, -2.605373, -0.778123, 1.570796, 2.139302],accel_mss,speed_ms,0,blend_radius_m)
  movel([0.561322, -1.324281, -2.608284, -0.779825, 1.570796, 2.132118],accel_mss,speed_ms,0,blend_radius_m)
  movel([0.552872, -1.319691, -2.611152, -0.781547, 1.570796, 2.123668],accel_mss,speed_ms,0,blend_radius_m)
  movel([0.548266, -1.317762, -2.612348, -0.782279, 1.570796, 2.119062],accel_mss,speed_ms,0,blend_radius_m)
  movel([0.543456, -1.316269, -2.613271, -0.782849, 1.570796, 2.114252],accel_mss,speed_ms,0,blend_radius_m)
  movel([0.538497, -1.315354, -2.613836, -0.783200, 1.570796, 2.109293],accel_mss,speed_ms,0,blend_radius_m)
  movel([0.533436, -1.315155, -2.613958, -0.783276, 1.570796, 2.104233],accel_mss,speed_ms,0,blend_radius_m)
  movel([0.528330, -1.315804, -2.613558, -0.783027, 1.570796, 2.099126],accel_mss,speed_ms,0,blend_radius_m)
  movel([0.523241, -1.317432, -2.612552, -0.782404, 1.570796, 2.094037],accel_mss,speed_ms,0,blend_radius_m)
  movel([0.520723, -1.318650, -2.611798, -0.781941, 1.570796, 2.091519],accel_mss,speed_ms,0,blend_radius_m)
  movel([0.518232, -1.320159, -2.610860, -0.781370, 1.570796, 2.089028],accel_mss,speed_ms,0,blend_radius_m)
  movel([0.515777, -1.321970, -2.609731, -0.780688, 1.570796, 2.086573],accel_mss,speed_ms,0,blend_radius_m)
  movel([0.513367, -1.324097, -2.608399, -0.779893, 1.570796, 2.084163],accel_mss,speed_ms,0,blend_radius_m)
  movel([0.511012, -1.326553, -2.606854, -0.778983, 1.570796, 2.081808],accel_mss,speed_ms,0,blend_radius_m)
  movel([0.508715, -1.329347, -2.605085, -0.777956, 1.570796, 2.079511],accel_mss,speed_ms,0,blend_radius_m)
  movel([0.504344, -1.336005, -2.600830, -0.775555, 1.570796, 2.075140],accel_mss,speed_ms,0,blend_radius_m)
  movel([0.503052, -1.339278, -2.598716, -0.774396, 1.570796, 2.073849],accel_mss,speed_ms,0,blend_radius_m)
  movel([0.502373, -1.342549, -2.596588, -0.773252, 1.570796, 2.073169],accel_mss,speed_ms,0,blend_radius_m)
  movel([0.502353, -1.345782, -2.594471, -0.772136, 1.570796, 2.073149],accel_mss,speed_ms,0,blend_radius_m)
  movel([0.503033, -1.348947, -2.592384, -0.771058, 1.570796, 2.073829],accel_mss,speed_ms,0,blend_radius_m)
  movel([0.506662, -1.344951, -2.595016, -0.772422, 1.570796, 2.077459],accel_mss,speed_ms,0,blend_radius_m)
  movel([0.510517, -1.341303, -2.597400, -0.773686, 1.570796, 2.081314],accel_mss,speed_ms,0,blend_radius_m)
  movel([0.514553, -1.338023, -2.599528, -0.774838, 1.570796, 2.085349],accel_mss,speed_ms,0,blend_radius_m)
  movel([0.518729, -1.335129, -2.601393, -0.775867, 1.570796, 2.089526],accel_mss,speed_ms,0,blend_radius_m)
  movel([0.523004, -1.332636, -2.602991, -0.776763, 1.570796, 2.093801],accel_mss,speed_ms,0,blend_radius_m)
  movel([0.527329, -1.330563, -2.604313, -0.777513, 1.570796, 2.098125],accel_mss,speed_ms,0,blend_radius_m)
  movel([0.531664, -1.328924, -2.605354, -0.778111, 1.570796, 2.102460],accel_mss,speed_ms,0,blend_radius_m)
  movel([0.535960, -1.327735, -2.606106, -0.778547, 1.570796, 2.106756],accel_mss,speed_ms,0,blend_radius_m)
  movel([0.540176, -1.327006, -2.606567, -0.778815, 1.570796, 2.110972],accel_mss,speed_ms,0,blend_radius_m)
  movel([0.544263, -1.326753, -2.606727, -0.778909, 1.570796, 2.115059],accel_mss,speed_ms,0,blend_radius_m)
  movel([0.548180, -1.326984, -2.606582, -0.778824, 1.570796, 2.118977],accel_mss,speed_ms,0,blend_radius_m)
  movel([0.551882, -1.327703, -2.606127, -0.778559, 1.570796, 2.122679],accel_mss,speed_ms,0,blend_radius_m)
  movel([0.555326, -1.328922, -2.605355, -0.778112, 1.570796, 2.126122],accel_mss,speed_ms,0,blend_radius_m)
  movel([0.558473, -1.330642, -2.604262, -0.777485, 1.570796, 2.129269],accel_mss,speed_ms,0,blend_radius_m)
  movel([0.561278, -1.332868, -2.602842, -0.776679, 1.570796, 2.132074],accel_mss,speed_ms,0,blend_radius_m)
  movel([0.563708, -1.335599, -2.601091, -0.775699, 1.570796, 2.134504],accel_mss,speed_ms,0,blend_radius_m)
  movel([0.565340, -1.338157, -2.599441, -0.774791, 1.570796, 2.136136],accel_mss,speed_ms,0,blend_radius_m)
  movel([0.566561, -1.340877, -2.597677, -0.773835, 1.570796, 2.137357],accel_mss,speed_ms,0,blend_radius_m)
  movel([0.567395, -1.343730, -2.595816, -0.772843, 1.570796, 2.138191],accel_mss,speed_ms,0,blend_radius_m)
  movel([0.567862, -1.346693, -2.593872, -0.771824, 1.570796, 2.138658],accel_mss,speed_ms,0,blend_radius_m)
  movel([0.567770, -1.352854, -2.589789, -0.769746, 1.570796, 2.138566],accel_mss,speed_ms,0,blend_radius_m)
  movel([0.566448, -1.359182, -2.585542, -0.767666, 1.570796, 2.137245],accel_mss,speed_ms,0,blend_radius_m)
  movel([0.564051, -1.365500, -2.581244, -0.765645, 1.570796, 2.134848],accel_mss,speed_ms,0,blend_radius_m)
  movel([0.560730, -1.371656, -2.577003, -0.763730, 1.570796, 2.131526],accel_mss,speed_ms,0,blend_radius_m)
  movel([0.556628, -1.377496, -2.572930, -0.761963, 1.570796, 2.127425],accel_mss,speed_ms,0,blend_radius_m)
  movel([0.551876, -1.382876, -2.569134, -0.760379, 1.570796, 2.122672],accel_mss,speed_ms,0,blend_radius_m)
  movel([0.546600, -1.387662, -2.565723, -0.759004, 1.570796, 2.117396],accel_mss,speed_ms,0,blend_radius_m)
  movel([0.540916, -1.391721, -2.562803, -0.757864, 1.570796, 2.111712],accel_mss,speed_ms,0,blend_radius_m)
  movel([0.534936, -1.394924, -2.560483, -0.756982, 1.570796, 2.105732],accel_mss,speed_ms,0,blend_radius_m)
  movel([0.531867, -1.396162, -2.559582, -0.756645, 1.570796, 2.102663],accel_mss,speed_ms,0,blend_radius_m)
  movel([0.528763, -1.397138, -2.558870, -0.756381, 1.570796, 2.099559],accel_mss,speed_ms,0,blend_radius_m)
  movel([0.525637, -1.397831, -2.558364, -0.756194, 1.570796, 2.096433],accel_mss,speed_ms,0,blend_radius_m)
  movel([0.522494, -1.398229, -2.558073, -0.756087, 1.570796, 2.093291],accel_mss,speed_ms,0,blend_radius_m)
  movel([0.519351, -1.398315, -2.558010, -0.756064, 1.570796, 2.090148],accel_mss,speed_ms,0,blend_radius_m)
  movel([0.516222, -1.398067, -2.558192, -0.756131, 1.570796, 2.087018],accel_mss,speed_ms,0,blend_radius_m)
  movel([0.513111, -1.397469, -2.558629, -0.756291, 1.570796, 2.083907],accel_mss,speed_ms,0,blend_radius_m)
  movel([0.510032, -1.396501, -2.559335, -0.756553, 1.570796, 2.080829],accel_mss,speed_ms,0,blend_radius_m)
  movel([0.506997, -1.395146, -2.560322, -0.756921, 1.570796, 2.077793],accel_mss,speed_ms,0,blend_radius_m)
  movel([0.504015, -1.393382, -2.561602, -0.757405, 1.570796, 2.074812],accel_mss,speed_ms,0,blend_radius_m)
  movel([0.501981, -1.391526, -2.562944, -0.757919, 1.570796, 2.072778],accel_mss,speed_ms,0,blend_radius_m)
  movel([0.497007, -1.385771, -2.567075, -0.759543, 1.570796, 2.067804],accel_mss,speed_ms,0,blend_radius_m)
  movel([0.493932, -1.381330, -2.570229, -0.760830, 1.570796, 2.064729],accel_mss,speed_ms,0,blend_radius_m)
  movel([0.490743, -1.375781, -2.574131, -0.762477, 1.570796, 2.061539],accel_mss,speed_ms,0,blend_radius_m)
  movel([0.487651, -1.369061, -2.578798, -0.764531, 1.570796, 2.058447],accel_mss,speed_ms,0,blend_radius_m)
  movel([0.484874, -1.361095, -2.584246, -0.767048, 1.570796, 2.055670],accel_mss,speed_ms,0,blend_radius_m)
  movel([0.483484, -1.355150, -2.588254, -0.768985, 1.570796, 2.054280],accel_mss,speed_ms,0,blend_radius_m)
  movel([0.482825, -1.349421, -2.592071, -0.770898, 1.570796, 2.053622],accel_mss,speed_ms,0,blend_radius_m)
  movel([0.482824, -1.343923, -2.595690, -0.772776, 1.570796, 2.053620],accel_mss,speed_ms,0,blend_radius_m)
  movel([0.483398, -1.338680, -2.599103, -0.774606, 1.570796, 2.054194],accel_mss,speed_ms,0,blend_radius_m)
  movel([0.484471, -1.333708, -2.602304, -0.776376, 1.570796, 2.055267],accel_mss,speed_ms,0,blend_radius_m)
  movel([0.485948, -1.329034, -2.605284, -0.778071, 1.570796, 2.056744],accel_mss,speed_ms,0,blend_radius_m)
  movel([0.487747, -1.324683, -2.608031, -0.779675, 1.570796, 2.058543],accel_mss,speed_ms,0,blend_radius_m)
  movel([0.489769, -1.320681, -2.610535, -0.781173, 1.570796, 2.060565],accel_mss,speed_ms,0,blend_radius_m)
  movel([0.494114, -1.313830, -2.614773, -0.783786, 1.570796, 2.064911],accel_mss,speed_ms,0,blend_radius_m)
  movel([0.498202, -1.308697, -2.617907, -0.785785, 1.570796, 2.068999],accel_mss,speed_ms,0,blend_radius_m)
  movel([0.501237, -1.305484, -2.619852, -0.787054, 1.570796, 2.072033],accel_mss,speed_ms,0,blend_radius_m)
  movel([0.502421, -1.304375, -2.620519, -0.787495, 1.570796, 2.073218],accel_mss,speed_ms,0,blend_radius_m)
  movel([0.508263, -1.299473, -2.623453, -0.789463, 1.570796, 2.079059],accel_mss,speed_ms,0,blend_radius_m)
  movel([0.514068, -1.295345, -2.625899, -0.791145, 1.570796, 2.084865],accel_mss,speed_ms,0,blend_radius_m)
  movel([0.519787, -1.291944, -2.627898, -0.792547, 1.570796, 2.090584],accel_mss,speed_ms,0,blend_radius_m)
  movel([0.525379, -1.289225, -2.629485, -0.793678, 1.570796, 2.096176],accel_mss,speed_ms,0,blend_radius_m)
  movel([0.530798, -1.287133, -2.630700, -0.794555, 1.570796, 2.101594],accel_mss,speed_ms,0,blend_radius_m)
  movel([0.536001, -1.285615, -2.631578, -0.795195, 1.570796, 2.106797],accel_mss,speed_ms,0,blend_radius_m)
  movel([0.540955, -1.284607, -2.632160, -0.795622, 1.570796, 2.111752],accel_mss,speed_ms,0,blend_radius_m)
  movel([0.545619, -1.284050, -2.632481, -0.795858, 1.570796, 2.116415],accel_mss,speed_ms,0,blend_radius_m)
  movel([0.553945, -1.284016, -2.632500, -0.795872, 1.570796, 2.124741],accel_mss,speed_ms,0,blend_radius_m)
  movel([0.560743, -1.284965, -2.631954, -0.795470, 1.570796, 2.131539],accel_mss,speed_ms,0,blend_radius_m)
  movel([0.565796, -1.286340, -2.631160, -0.794889, 1.570796, 2.136592],accel_mss,speed_ms,0,blend_radius_m)
  movel([0.568914, -1.287574, -2.630445, -0.794370, 1.570796, 2.139710],accel_mss,speed_ms,0,blend_radius_m)
  movel([0.576341, -1.290443, -2.628776, -0.793171, 1.570796, 2.147137],accel_mss,speed_ms,0,blend_radius_m)
  movel([0.583895, -1.294245, -2.626547, -0.791597, 1.570796, 2.154691],accel_mss,speed_ms,0,blend_radius_m)
  movel([0.591384, -1.298355, -2.624117, -0.789916, 1.570796, 2.162180],accel_mss,speed_ms,0,blend_radius_m)
  movel([0.598645, -1.302153, -2.621853, -0.788383, 1.570796, 2.169441],accel_mss,speed_ms,0,blend_radius_m)
  movel([0.605543, -1.305014, -2.620135, -0.787240, 1.570796, 2.176339],accel_mss,speed_ms,0,blend_radius_m)
  movel([0.608818, -1.305896, -2.619603, -0.786890, 1.570796, 2.179614],accel_mss,speed_ms,0,blend_radius_m)
  movel([0.611960, -1.306308, -2.619354, -0.786727, 1.570796, 2.182756],accel_mss,speed_ms,0,blend_radius_m)
  movel([0.614956, -1.306168, -2.619439, -0.786782, 1.570796, 2.185753],accel_mss,speed_ms,0,blend_radius_m)
  movel([0.617798, -1.305393, -2.619907, -0.787090, 1.570796, 2.188595],accel_mss,speed_ms,0,blend_radius_m)
  movel([0.620474, -1.303901, -2.620804, -0.787684, 1.570796, 2.191271],accel_mss,speed_ms,0,blend_radius_m)
  movel([0.622972, -1.301603, -2.622182, -0.788604, 1.570796, 2.193768],accel_mss,speed_ms,0,blend_radius_m)
  movel([0.624521, -1.299621, -2.623365, -0.789403, 1.570796, 2.195317],accel_mss,speed_ms,0,blend_radius_m)
  movel([0.625698, -1.297638, -2.624543, -0.790208, 1.570796, 2.196494],accel_mss,speed_ms,0,blend_radius_m)
  movel([0.627084, -1.293678, -2.626881, -0.791830, 1.570796, 2.197881],accel_mss,speed_ms,0,blend_radius_m)
  movel([0.627416, -1.289738, -2.629187, -0.793464, 1.570796, 2.198213],accel_mss,speed_ms,0,blend_radius_m)
  movel([0.626972, -1.285848, -2.631444, -0.795097, 1.570796, 2.197768],accel_mss,speed_ms,0,blend_radius_m)
  movel([0.624932, -1.278300, -2.635769, -0.798320, 1.570796, 2.195728],accel_mss,speed_ms,0,blend_radius_m)
  movel([0.623931, -1.274685, -2.637816, -0.799888, 1.570796, 2.194728],accel_mss,speed_ms,0,blend_radius_m)
  movel([0.623355, -1.271197, -2.639775, -0.801417, 1.570796, 2.194152],accel_mss,speed_ms,0,blend_radius_m)
  movel([0.623591, -1.265467, -2.642960, -0.803962, 1.570796, 2.194388],accel_mss,speed_ms,0,blend_radius_m)
  movel([0.624822, -1.258164, -2.646962, -0.807263, 1.570796, 2.195618],accel_mss,speed_ms,0,blend_radius_m)
  movel([0.626768, -1.250595, -2.651041, -0.810753, 1.570796, 2.197564],accel_mss,speed_ms,0,blend_radius_m)
  movel([0.629130, -1.244133, -2.654469, -0.813787, 1.570796, 2.199927],accel_mss,speed_ms,0,blend_radius_m)
  movel([0.631408, -1.240121, -2.656572, -0.815696, 1.570796, 2.202204],accel_mss,speed_ms,0,blend_radius_m)
  movel([0.634597, -1.235244, -2.659104, -0.818041, 1.570796, 2.205393],accel_mss,speed_ms,0,blend_radius_m)
  movel([0.637598, -1.230585, -2.661496, -0.820307, 1.570796, 2.208394],accel_mss,speed_ms,0,blend_radius_m)
  movel([0.639286, -1.227254, -2.663191, -0.821943, 1.570796, 2.210082],accel_mss,speed_ms,0,blend_radius_m)
  movel([0.639664, -1.223919, -2.664876, -0.823595, 1.570796, 2.210460],accel_mss,speed_ms,0,blend_radius_m)
  movel([0.639450, -1.220151, -2.666763, -0.825475, 1.570796, 2.210247],accel_mss,speed_ms,0,blend_radius_m)
  movel([0.639270, -1.215923, -2.668862, -0.827604, 1.570796, 2.210066],accel_mss,speed_ms,0,blend_radius_m)
  movel([0.639773, -1.211195, -2.671185, -0.830009, 1.570796, 2.210569],accel_mss,speed_ms,0,blend_radius_m)
  movel([0.640733, -1.208251, -2.672619, -0.831519, 1.570796, 2.211529],accel_mss,speed_ms,0,blend_radius_m)
  speed_ms = 0.003
  movel([0.640733, -1.200996, -2.669029, -0.842364, 1.570796, 2.211529],accel_mss,speed_ms,0,blend_radius_m)
  speed_ms = 0.03
  movel([0.640733, -1.173424, -2.654409, -0.884556, 1.570796, 2.211529],accel_mss,speed_ms,0,blend_radius_m)
  #M_RunCode9
  movel([0.485052, -1.296681, -2.588792, -0.826916, 1.570796, 2.055849],accel_mss,speed_ms,0,blend_radius_m)
  #M_RunCode3
  movel([0.485052, -1.322750, -2.601783, -0.787856, 1.570796, 2.055849],accel_mss,speed_ms,0,blend_radius_m)
  speed_ms = 0.003
  movel([0.485052, -1.329545, -2.604960, -0.777884, 1.570796, 2.055849],accel_mss,speed_ms,0,blend_radius_m)
  speed_ms = 0.007
  movel([0.477144, -1.327685, -2.606138, -0.778566, 1.570796, 2.047940],accel_mss,speed_ms,0,blend_radius_m)
  movel([0.469118, -1.326870, -2.606653, -0.778865, 1.570796, 2.039914],accel_mss,speed_ms,0,blend_radius_m)
  movel([0.461080, -1.326977, -2.606586, -0.778826, 1.570796, 2.031877],accel_mss,speed_ms,0,blend_radius_m)
  movel([0.453131, -1.327874, -2.606019, -0.778496, 1.570796, 2.023928],accel_mss,speed_ms,0,blend_radius_m)
  movel([0.445372, -1.329430, -2.605033, -0.777926, 1.570796, 2.016168],accel_mss,speed_ms,0,blend_radius_m)
  movel([0.437898, -1.331510, -2.603710, -0.777170, 1.570796, 2.008694],accel_mss,speed_ms,0,blend_radius_m)
  movel([0.430791, -1.333985, -2.602127, -0.776277, 1.570796, 2.001587],accel_mss,speed_ms,0,blend_radius_m)
  movel([0.424140, -1.336718, -2.600370, -0.775301, 1.570796, 1.994937],accel_mss,speed_ms,0,blend_radius_m)
  movel([0.418019, -1.339583, -2.598518, -0.774288, 1.570796, 1.988816],accel_mss,speed_ms,0,blend_radius_m)
  movel([0.412504, -1.342453, -2.596651, -0.773286, 1.570796, 1.983300],accel_mss,speed_ms,0,blend_radius_m)
  movel([0.403562, -1.347709, -2.593202, -0.771478, 1.570796, 1.974358],accel_mss,speed_ms,0,blend_radius_m)
  movel([0.397826, -1.351539, -2.590665, -0.770185, 1.570796, 1.968622],accel_mss,speed_ms,0,blend_radius_m)
  movel([0.395803, -1.353016, -2.589681, -0.769692, 1.570796, 1.966599],accel_mss,speed_ms,0,blend_radius_m)
  movel([0.392530, -1.355264, -2.588178, -0.768947, 1.570796, 1.963326],accel_mss,speed_ms,0,blend_radius_m)
  movel([0.384260, -1.361692, -2.583841, -0.766856, 1.570796, 1.955056],accel_mss,speed_ms,0,blend_radius_m)
  movel([0.378988, -1.366313, -2.580687, -0.765389, 1.570796, 1.949785],accel_mss,speed_ms,0,blend_radius_m)
  movel([0.373353, -1.371774, -2.576921, -0.763694, 1.570796, 1.944149],accel_mss,speed_ms,0,blend_radius_m)
  movel([0.367647, -1.377996, -2.572579, -0.761814, 1.570796, 1.938443],accel_mss,speed_ms,0,blend_radius_m)
  movel([0.362155, -1.384903, -2.567693, -0.759792, 1.570796, 1.932952],accel_mss,speed_ms,0,blend_radius_m)
  movel([0.357157, -1.392407, -2.562307, -0.757674, 1.570796, 1.927953],accel_mss,speed_ms,0,blend_radius_m)
  movel([0.352917, -1.400432, -2.556457, -0.755499, 1.570796, 1.923713],accel_mss,speed_ms,0,blend_radius_m)
  movel([0.351159, -1.404616, -2.553370, -0.754403, 1.570796, 1.921955],accel_mss,speed_ms,0,blend_radius_m)
  movel([0.349687, -1.408900, -2.550182, -0.753307, 1.570796, 1.920483],accel_mss,speed_ms,0,blend_radius_m)
  movel([0.348525, -1.413278, -2.546896, -0.752215, 1.570796, 1.919322],accel_mss,speed_ms,0,blend_radius_m)
  movel([0.347704, -1.417741, -2.543517, -0.751131, 1.570796, 1.918501],accel_mss,speed_ms,0,blend_radius_m)
  movel([0.347253, -1.422282, -2.540048, -0.750059, 1.570796, 1.918049],accel_mss,speed_ms,0,blend_radius_m)
  movel([0.347196, -1.426896, -2.536492, -0.749001, 1.570796, 1.917992],accel_mss,speed_ms,0,blend_radius_m)
  movel([0.347560, -1.431575, -2.532853, -0.747961, 1.570796, 1.918357],accel_mss,speed_ms,0,blend_radius_m)
  movel([0.348366, -1.436315, -2.529133, -0.746941, 1.570796, 1.919163],accel_mss,speed_ms,0,blend_radius_m)
  movel([0.349641, -1.441115, -2.525331, -0.745943, 1.570796, 1.920437],accel_mss,speed_ms,0,blend_radius_m)
  movel([0.351404, -1.445968, -2.521452, -0.744969, 1.570796, 1.922200],accel_mss,speed_ms,0,blend_radius_m)
  movel([0.353676, -1.450876, -2.517492, -0.744021, 1.570796, 1.924472],accel_mss,speed_ms,0,blend_radius_m)
  movel([0.356480, -1.455837, -2.513451, -0.743100, 1.570796, 1.927277],accel_mss,speed_ms,0,blend_radius_m)
  movel([0.356730, -1.456203, -2.513152, -0.743034, 1.570796, 1.927526],accel_mss,speed_ms,0,blend_radius_m)
  movel([0.360297, -1.460589, -2.509546, -0.742254, 1.570796, 1.931093],accel_mss,speed_ms,0,blend_radius_m)
  movel([0.363954, -1.464426, -2.506367, -0.741596, 1.570796, 1.934750],accel_mss,speed_ms,0,blend_radius_m)
  movel([0.367690, -1.467746, -2.503599, -0.741045, 1.570796, 1.938487],accel_mss,speed_ms,0,blend_radius_m)
  movel([0.371495, -1.470582, -2.501219, -0.740588, 1.570796, 1.942291],accel_mss,speed_ms,0,blend_radius_m)
  movel([0.375360, -1.472965, -2.499211, -0.740213, 1.570796, 1.946156],accel_mss,speed_ms,0,blend_radius_m)
  movel([0.379274, -1.474924, -2.497553, -0.739912, 1.570796, 1.950070],accel_mss,speed_ms,0,blend_radius_m)
  movel([0.383222, -1.476489, -2.496224, -0.739676, 1.570796, 1.954018],accel_mss,speed_ms,0,blend_radius_m)
  movel([0.387196, -1.477686, -2.495205, -0.739498, 1.570796, 1.957993],accel_mss,speed_ms,0,blend_radius_m)
  movel([0.391186, -1.478544, -2.494474, -0.739371, 1.570796, 1.961982],accel_mss,speed_ms,0,blend_radius_m)
  movel([0.395180, -1.479084, -2.494012, -0.739292, 1.570796, 1.965976],accel_mss,speed_ms,0,blend_radius_m)
  movel([0.399163, -1.479337, -2.493797, -0.739255, 1.570796, 1.969959],accel_mss,speed_ms,0,blend_radius_m)
  movel([0.403126, -1.479323, -2.493808, -0.739257, 1.570796, 1.973922],accel_mss,speed_ms,0,blend_radius_m)
  movel([0.410930, -1.478603, -2.494424, -0.739363, 1.570796, 1.981727],accel_mss,speed_ms,0,blend_radius_m)
  movel([0.418492, -1.477116, -2.495691, -0.739582, 1.570796, 1.989288],accel_mss,speed_ms,0,blend_radius_m)
  movel([0.425688, -1.475057, -2.497440, -0.739892, 1.570796, 1.996484],accel_mss,speed_ms,0,blend_radius_m)
  movel([0.432396, -1.472618, -2.499504, -0.740267, 1.570796, 2.003192],accel_mss,speed_ms,0,blend_radius_m)
  movel([0.438480, -1.469995, -2.501712, -0.740681, 1.570796, 2.009276],accel_mss,speed_ms,0,blend_radius_m)
  movel([0.443800, -1.467387, -2.503899, -0.741104, 1.570796, 2.014596],accel_mss,speed_ms,0,blend_radius_m)
  movel([0.451548, -1.463028, -2.507528, -0.741833, 1.570796, 2.022345],accel_mss,speed_ms,0,blend_radius_m)
  movel([0.454404, -1.461200, -2.509042, -0.742148, 1.570796, 2.025201],accel_mss,speed_ms,0,blend_radius_m)
  movel([0.456159, -1.460139, -2.509917, -0.742333, 1.570796, 2.026955],accel_mss,speed_ms,0,blend_radius_m)
  movel([0.460906, -1.457017, -2.512485, -0.742887, 1.570796, 2.031703],accel_mss,speed_ms,0,blend_radius_m)
  movel([0.467900, -1.451902, -2.516659, -0.743828, 1.570796, 2.038696],accel_mss,speed_ms,0,blend_radius_m)
  movel([0.476405, -1.444846, -2.522352, -0.745191, 1.570796, 2.047202],accel_mss,speed_ms,0,blend_radius_m)
  movel([0.480996, -1.440597, -2.525743, -0.746049, 1.570796, 2.051793],accel_mss,speed_ms,0,blend_radius_m)
  movel([0.485693, -1.435867, -2.529486, -0.747036, 1.570796, 2.056489],accel_mss,speed_ms,0,blend_radius_m)
  movel([0.490400, -1.430657, -2.533569, -0.748162, 1.570796, 2.061196],accel_mss,speed_ms,0,blend_radius_m)
  movel([0.495024, -1.424959, -2.537989, -0.749441, 1.570796, 2.065820],accel_mss,speed_ms,0,blend_radius_m)
  movel([0.499466, -1.418769, -2.542734, -0.750886, 1.570796, 2.070262],accel_mss,speed_ms,0,blend_radius_m)
  movel([0.503628, -1.412078, -2.547799, -0.752512, 1.570796, 2.074424],accel_mss,speed_ms,0,blend_radius_m)
  movel([0.507405, -1.404881, -2.553174, -0.754334, 1.570796, 2.078201],accel_mss,speed_ms,0,blend_radius_m)
  movel([0.510691, -1.397163, -2.558852, -0.756374, 1.570796, 2.081487],accel_mss,speed_ms,0,blend_radius_m)
  speed_ms = 0.003
  movel([0.510691, -1.390712, -2.555900, -0.765777, 1.570796, 2.081487],accel_mss,speed_ms,0,blend_radius_m)
  speed_ms = 0.03
  movel([0.510691, -1.365852, -2.543800, -0.802737, 1.570796, 2.081487],accel_mss,speed_ms,0,blend_radius_m)
  #M_RunCode9
  movel([0.478180, -1.358037, -2.549202, -0.805149, 1.570796, 2.048976],accel_mss,speed_ms,0,blend_radius_m)
  #M_RunCode3
